screen "Lists" 1920x1080, template "Tpl"
   TextField "frm_1" at 16,154 size 1888x84; Text 'Text'
   TextField "txt_1" at 28,158 size 400x28; Text 'POSTAVKE (dok sustav stoji)'
   TextField "txt_2" at 28,194 size 160x34; Text 'Redoslijed'
   SymbolicIOField "sym_1" at 188,194 size 330x34; TextOff '0'; TextOn '1'; TextList "TL_Order"
      ProcessValue <- "CfgOrderMode"
   TextField "txt_3" at 560,194 size 290x34; Text 'SEMI: transfer po koraku'
   SymbolicIOField "sym_2" at 850,194 size 110x34; TextOff '0'; TextOn '1'; TextList "TL_YesNo"
      ProcessValue <- "CfgSemiPerTransfer"
   TextField "txt_4" at 1000,194 size 180x34; Text 'Ravnoteža'
   SymbolicIOField "sym_3" at 1180,194 size 260x34; TextOff '0'; TextOn '1'; TextList "TL_BalMode"
      ProcessValue <- "CfgBalMode"
   TextField "txt_5" at 1480,194 size 80x34; Text 'Istovar'
   IOField "io_1" at 1560,194 size 60x34; FormatPattern 99
      ProcessValue <- "UTotal"
   TextField "txt_6" at 1640,194 size 80x34; Text 'Ukrcaj'
   IOField "io_2" at 1720,194 size 60x34; FormatPattern 99
      ProcessValue <- "LTotal"
   TextField "txt_7" at 16,252 size 466x28; Text 'LISTA ZA ISTOVAR (DB20) 1-24'
   TextField "txt_8" at 16,286 size 46x27; Text '1'
   IOField "io_3" at 68,286 size 90x27; FormatPattern 999
      ProcessValue <- "UList_01"
   SymbolicIOField "sym_4" at 164,286 size 150x27; TextOff '0'; TextOn '1'; TextList "TL_ListSt"
      ProcessValue <- "UState_01"
   TextField "txt_9" at 16,316 size 46x27; Text '2'
   IOField "io_4" at 68,316 size 90x27; FormatPattern 999
      ProcessValue <- "UList_02"
   SymbolicIOField "sym_5" at 164,316 size 150x27; TextOff '0'; TextOn '1'; TextList "TL_ListSt"
      ProcessValue <- "UState_02"
   TextField "txt_10" at 16,346 size 46x27; Text '3'
   IOField "io_5" at 68,346 size 90x27; FormatPattern 999
      ProcessValue <- "UList_03"
   SymbolicIOField "sym_6" at 164,346 size 150x27; TextOff '0'; TextOn '1'; TextList "TL_ListSt"
      ProcessValue <- "UState_03"
   TextField "txt_11" at 16,376 size 46x27; Text '4'
   IOField "io_6" at 68,376 size 90x27; FormatPattern 999
      ProcessValue <- "UList_04"
   SymbolicIOField "sym_7" at 164,376 size 150x27; TextOff '0'; TextOn '1'; TextList "TL_ListSt"
      ProcessValue <- "UState_04"
   TextField "txt_12" at 16,406 size 46x27; Text '5'
   IOField "io_7" at 68,406 size 90x27; FormatPattern 999
      ProcessValue <- "UList_05"
   SymbolicIOField "sym_8" at 164,406 size 150x27; TextOff '0'; TextOn '1'; TextList "TL_ListSt"
      ProcessValue <- "UState_05"
   TextField "txt_13" at 16,436 size 46x27; Text '6'
   IOField "io_8" at 68,436 size 90x27; FormatPattern 999
      ProcessValue <- "UList_06"
   SymbolicIOField "sym_9" at 164,436 size 150x27; TextOff '0'; TextOn '1'; TextList "TL_ListSt"
      ProcessValue <- "UState_06"
   TextField "txt_14" at 16,466 size 46x27; Text '7'
   IOField "io_9" at 68,466 size 90x27; FormatPattern 999
      ProcessValue <- "UList_07"
   SymbolicIOField "sym_10" at 164,466 size 150x27; TextOff '0'; TextOn '1'; TextList "TL_ListSt"
      ProcessValue <- "UState_07"
   TextField "txt_15" at 16,496 size 46x27; Text '8'
   IOField "io_10" at 68,496 size 90x27; FormatPattern 999
      ProcessValue <- "UList_08"
   SymbolicIOField "sym_11" at 164,496 size 150x27; TextOff '0'; TextOn '1'; TextList "TL_ListSt"
      ProcessValue <- "UState_08"
   TextField "txt_16" at 16,526 size 46x27; Text '9'
   IOField "io_11" at 68,526 size 90x27; FormatPattern 999
      ProcessValue <- "UList_09"
   SymbolicIOField "sym_12" at 164,526 size 150x27; TextOff '0'; TextOn '1'; TextList "TL_ListSt"
      ProcessValue <- "UState_09"
   TextField "txt_17" at 16,556 size 46x27; Text '10'
   IOField "io_12" at 68,556 size 90x27; FormatPattern 999
      ProcessValue <- "UList_10"
   SymbolicIOField "sym_13" at 164,556 size 150x27; TextOff '0'; TextOn '1'; TextList "TL_ListSt"
      ProcessValue <- "UState_10"
   TextField "txt_18" at 16,586 size 46x27; Text '11'
   IOField "io_13" at 68,586 size 90x27; FormatPattern 999
      ProcessValue <- "UList_11"
   SymbolicIOField "sym_14" at 164,586 size 150x27; TextOff '0'; TextOn '1'; TextList "TL_ListSt"
      ProcessValue <- "UState_11"
   TextField "txt_19" at 16,616 size 46x27; Text '12'
   IOField "io_14" at 68,616 size 90x27; FormatPattern 999
      ProcessValue <- "UList_12"
   SymbolicIOField "sym_15" at 164,616 size 150x27; TextOff '0'; TextOn '1'; TextList "TL_ListSt"
      ProcessValue <- "UState_12"
   TextField "txt_20" at 16,646 size 46x27; Text '13'
   IOField "io_15" at 68,646 size 90x27; FormatPattern 999
      ProcessValue <- "UList_13"
   SymbolicIOField "sym_16" at 164,646 size 150x27; TextOff '0'; TextOn '1'; TextList "TL_ListSt"
      ProcessValue <- "UState_13"
   TextField "txt_21" at 16,676 size 46x27; Text '14'
   IOField "io_16" at 68,676 size 90x27; FormatPattern 999
      ProcessValue <- "UList_14"
   SymbolicIOField "sym_17" at 164,676 size 150x27; TextOff '0'; TextOn '1'; TextList "TL_ListSt"
      ProcessValue <- "UState_14"
   TextField "txt_22" at 16,706 size 46x27; Text '15'
   IOField "io_17" at 68,706 size 90x27; FormatPattern 999
      ProcessValue <- "UList_15"
   SymbolicIOField "sym_18" at 164,706 size 150x27; TextOff '0'; TextOn '1'; TextList "TL_ListSt"
      ProcessValue <- "UState_15"
   TextField "txt_23" at 16,736 size 46x27; Text '16'
   IOField "io_18" at 68,736 size 90x27; FormatPattern 999
      ProcessValue <- "UList_16"
   SymbolicIOField "sym_19" at 164,736 size 150x27; TextOff '0'; TextOn '1'; TextList "TL_ListSt"
      ProcessValue <- "UState_16"
   TextField "txt_24" at 16,766 size 46x27; Text '17'
   IOField "io_19" at 68,766 size 90x27; FormatPattern 999
      ProcessValue <- "UList_17"
   SymbolicIOField "sym_20" at 164,766 size 150x27; TextOff '0'; TextOn '1'; TextList "TL_ListSt"
      ProcessValue <- "UState_17"
   TextField "txt_25" at 16,796 size 46x27; Text '18'
   IOField "io_20" at 68,796 size 90x27; FormatPattern 999
      ProcessValue <- "UList_18"
   SymbolicIOField "sym_21" at 164,796 size 150x27; TextOff '0'; TextOn '1'; TextList "TL_ListSt"
      ProcessValue <- "UState_18"
   TextField "txt_26" at 16,826 size 46x27; Text '19'
   IOField "io_21" at 68,826 size 90x27; FormatPattern 999
      ProcessValue <- "UList_19"
   SymbolicIOField "sym_22" at 164,826 size 150x27; TextOff '0'; TextOn '1'; TextList "TL_ListSt"
      ProcessValue <- "UState_19"
   TextField "txt_27" at 16,856 size 46x27; Text '20'
   IOField "io_22" at 68,856 size 90x27; FormatPattern 999
      ProcessValue <- "UList_20"
   SymbolicIOField "sym_23" at 164,856 size 150x27; TextOff '0'; TextOn '1'; TextList "TL_ListSt"
      ProcessValue <- "UState_20"
   TextField "txt_28" at 16,886 size 46x27; Text '21'
   IOField "io_23" at 68,886 size 90x27; FormatPattern 999
      ProcessValue <- "UList_21"
   SymbolicIOField "sym_24" at 164,886 size 150x27; TextOff '0'; TextOn '1'; TextList "TL_ListSt"
      ProcessValue <- "UState_21"
   TextField "txt_29" at 16,916 size 46x27; Text '22'
   IOField "io_24" at 68,916 size 90x27; FormatPattern 999
      ProcessValue <- "UList_22"
   SymbolicIOField "sym_25" at 164,916 size 150x27; TextOff '0'; TextOn '1'; TextList "TL_ListSt"
      ProcessValue <- "UState_22"
   TextField "txt_30" at 16,946 size 46x27; Text '23'
   IOField "io_25" at 68,946 size 90x27; FormatPattern 999
      ProcessValue <- "UList_23"
   SymbolicIOField "sym_26" at 164,946 size 150x27; TextOff '0'; TextOn '1'; TextList "TL_ListSt"
      ProcessValue <- "UState_23"
   TextField "txt_31" at 16,976 size 46x27; Text '24'
   IOField "io_26" at 68,976 size 90x27; FormatPattern 999
      ProcessValue <- "UList_24"
   SymbolicIOField "sym_27" at 164,976 size 150x27; TextOff '0'; TextOn '1'; TextList "TL_ListSt"
      ProcessValue <- "UState_24"
   TextField "txt_32" at 490,252 size 466x28; Text 'LISTA ZA ISTOVAR 25-48'
   TextField "txt_33" at 490,286 size 46x27; Text '25'
   IOField "io_27" at 542,286 size 90x27; FormatPattern 999
      ProcessValue <- "UList_25"
   SymbolicIOField "sym_28" at 638,286 size 150x27; TextOff '0'; TextOn '1'; TextList "TL_ListSt"
      ProcessValue <- "UState_25"
   TextField "txt_34" at 490,316 size 46x27; Text '26'
   IOField "io_28" at 542,316 size 90x27; FormatPattern 999
      ProcessValue <- "UList_26"
   SymbolicIOField "sym_29" at 638,316 size 150x27; TextOff '0'; TextOn '1'; TextList "TL_ListSt"
      ProcessValue <- "UState_26"
   TextField "txt_35" at 490,346 size 46x27; Text '27'
   IOField "io_29" at 542,346 size 90x27; FormatPattern 999
      ProcessValue <- "UList_27"
   SymbolicIOField "sym_30" at 638,346 size 150x27; TextOff '0'; TextOn '1'; TextList "TL_ListSt"
      ProcessValue <- "UState_27"
   TextField "txt_36" at 490,376 size 46x27; Text '28'
   IOField "io_30" at 542,376 size 90x27; FormatPattern 999
      ProcessValue <- "UList_28"
   SymbolicIOField "sym_31" at 638,376 size 150x27; TextOff '0'; TextOn '1'; TextList "TL_ListSt"
      ProcessValue <- "UState_28"
   TextField "txt_37" at 490,406 size 46x27; Text '29'
   IOField "io_31" at 542,406 size 90x27; FormatPattern 999
      ProcessValue <- "UList_29"
   SymbolicIOField "sym_32" at 638,406 size 150x27; TextOff '0'; TextOn '1'; TextList "TL_ListSt"
      ProcessValue <- "UState_29"
   TextField "txt_38" at 490,436 size 46x27; Text '30'
   IOField "io_32" at 542,436 size 90x27; FormatPattern 999
      ProcessValue <- "UList_30"
   SymbolicIOField "sym_33" at 638,436 size 150x27; TextOff '0'; TextOn '1'; TextList "TL_ListSt"
      ProcessValue <- "UState_30"
   TextField "txt_39" at 490,466 size 46x27; Text '31'
   IOField "io_33" at 542,466 size 90x27; FormatPattern 999
      ProcessValue <- "UList_31"
   SymbolicIOField "sym_34" at 638,466 size 150x27; TextOff '0'; TextOn '1'; TextList "TL_ListSt"
      ProcessValue <- "UState_31"
   TextField "txt_40" at 490,496 size 46x27; Text '32'
   IOField "io_34" at 542,496 size 90x27; FormatPattern 999
      ProcessValue <- "UList_32"
   SymbolicIOField "sym_35" at 638,496 size 150x27; TextOff '0'; TextOn '1'; TextList "TL_ListSt"
      ProcessValue <- "UState_32"
   TextField "txt_41" at 490,526 size 46x27; Text '33'
   IOField "io_35" at 542,526 size 90x27; FormatPattern 999
      ProcessValue <- "UList_33"
   SymbolicIOField "sym_36" at 638,526 size 150x27; TextOff '0'; TextOn '1'; TextList "TL_ListSt"
      ProcessValue <- "UState_33"
   TextField "txt_42" at 490,556 size 46x27; Text '34'
   IOField "io_36" at 542,556 size 90x27; FormatPattern 999
      ProcessValue <- "UList_34"
   SymbolicIOField "sym_37" at 638,556 size 150x27; TextOff '0'; TextOn '1'; TextList "TL_ListSt"
      ProcessValue <- "UState_34"
   TextField "txt_43" at 490,586 size 46x27; Text '35'
   IOField "io_37" at 542,586 size 90x27; FormatPattern 999
      ProcessValue <- "UList_35"
   SymbolicIOField "sym_38" at 638,586 size 150x27; TextOff '0'; TextOn '1'; TextList "TL_ListSt"
      ProcessValue <- "UState_35"
   TextField "txt_44" at 490,616 size 46x27; Text '36'
   IOField "io_38" at 542,616 size 90x27; FormatPattern 999
      ProcessValue <- "UList_36"
   SymbolicIOField "sym_39" at 638,616 size 150x27; TextOff '0'; TextOn '1'; TextList "TL_ListSt"
      ProcessValue <- "UState_36"
   TextField "txt_45" at 490,646 size 46x27; Text '37'
   IOField "io_39" at 542,646 size 90x27; FormatPattern 999
      ProcessValue <- "UList_37"
   SymbolicIOField "sym_40" at 638,646 size 150x27; TextOff '0'; TextOn '1'; TextList "TL_ListSt"
      ProcessValue <- "UState_37"
   TextField "txt_46" at 490,676 size 46x27; Text '38'
   IOField "io_40" at 542,676 size 90x27; FormatPattern 999
      ProcessValue <- "UList_38"
   SymbolicIOField "sym_41" at 638,676 size 150x27; TextOff '0'; TextOn '1'; TextList "TL_ListSt"
      ProcessValue <- "UState_38"
   TextField "txt_47" at 490,706 size 46x27; Text '39'
   IOField "io_41" at 542,706 size 90x27; FormatPattern 999
      ProcessValue <- "UList_39"
   SymbolicIOField "sym_42" at 638,706 size 150x27; TextOff '0'; TextOn '1'; TextList "TL_ListSt"
      ProcessValue <- "UState_39"
   TextField "txt_48" at 490,736 size 46x27; Text '40'
   IOField "io_42" at 542,736 size 90x27; FormatPattern 999
      ProcessValue <- "UList_40"
   SymbolicIOField "sym_43" at 638,736 size 150x27; TextOff '0'; TextOn '1'; TextList "TL_ListSt"
      ProcessValue <- "UState_40"
   TextField "txt_49" at 490,766 size 46x27; Text '41'
   IOField "io_43" at 542,766 size 90x27; FormatPattern 999
      ProcessValue <- "UList_41"
   SymbolicIOField "sym_44" at 638,766 size 150x27; TextOff '0'; TextOn '1'; TextList "TL_ListSt"
      ProcessValue <- "UState_41"
   TextField "txt_50" at 490,796 size 46x27; Text '42'
   IOField "io_44" at 542,796 size 90x27; FormatPattern 999
      ProcessValue <- "UList_42"
   SymbolicIOField "sym_45" at 638,796 size 150x27; TextOff '0'; TextOn '1'; TextList "TL_ListSt"
      ProcessValue <- "UState_42"
   TextField "txt_51" at 490,826 size 46x27; Text '43'
   IOField "io_45" at 542,826 size 90x27; FormatPattern 999
      ProcessValue <- "UList_43"
   SymbolicIOField "sym_46" at 638,826 size 150x27; TextOff '0'; TextOn '1'; TextList "TL_ListSt"
      ProcessValue <- "UState_43"
   TextField "txt_52" at 490,856 size 46x27; Text '44'
   IOField "io_46" at 542,856 size 90x27; FormatPattern 999
      ProcessValue <- "UList_44"
   SymbolicIOField "sym_47" at 638,856 size 150x27; TextOff '0'; TextOn '1'; TextList "TL_ListSt"
      ProcessValue <- "UState_44"
   TextField "txt_53" at 490,886 size 46x27; Text '45'
   IOField "io_47" at 542,886 size 90x27; FormatPattern 999
      ProcessValue <- "UList_45"
   SymbolicIOField "sym_48" at 638,886 size 150x27; TextOff '0'; TextOn '1'; TextList "TL_ListSt"
      ProcessValue <- "UState_45"
   TextField "txt_54" at 490,916 size 46x27; Text '46'
   IOField "io_48" at 542,916 size 90x27; FormatPattern 999
      ProcessValue <- "UList_46"
   SymbolicIOField "sym_49" at 638,916 size 150x27; TextOff '0'; TextOn '1'; TextList "TL_ListSt"
      ProcessValue <- "UState_46"
   TextField "txt_55" at 490,946 size 46x27; Text '47'
   IOField "io_49" at 542,946 size 90x27; FormatPattern 999
      ProcessValue <- "UList_47"
   SymbolicIOField "sym_50" at 638,946 size 150x27; TextOff '0'; TextOn '1'; TextList "TL_ListSt"
      ProcessValue <- "UState_47"
   TextField "txt_56" at 490,976 size 46x27; Text '48'
   IOField "io_50" at 542,976 size 90x27; FormatPattern 999
      ProcessValue <- "UList_48"
   SymbolicIOField "sym_51" at 638,976 size 150x27; TextOff '0'; TextOn '1'; TextList "TL_ListSt"
      ProcessValue <- "UState_48"
   TextField "txt_57" at 964,252 size 466x28; Text 'LISTA ZA UKRCAJ (DB21) 1-24'
   TextField "txt_58" at 964,286 size 46x27; Text '1'
   IOField "io_51" at 1016,286 size 90x27; FormatPattern 999
      ProcessValue <- "LList_01"
   SymbolicIOField "sym_52" at 1112,286 size 150x27; TextOff '0'; TextOn '1'; TextList "TL_ListSt"
      ProcessValue <- "LState_01"
   TextField "txt_59" at 964,316 size 46x27; Text '2'
   IOField "io_52" at 1016,316 size 90x27; FormatPattern 999
      ProcessValue <- "LList_02"
   SymbolicIOField "sym_53" at 1112,316 size 150x27; TextOff '0'; TextOn '1'; TextList "TL_ListSt"
      ProcessValue <- "LState_02"
   TextField "txt_60" at 964,346 size 46x27; Text '3'
   IOField "io_53" at 1016,346 size 90x27; FormatPattern 999
      ProcessValue <- "LList_03"
   SymbolicIOField "sym_54" at 1112,346 size 150x27; TextOff '0'; TextOn '1'; TextList "TL_ListSt"
      ProcessValue <- "LState_03"
   TextField "txt_61" at 964,376 size 46x27; Text '4'
   IOField "io_54" at 1016,376 size 90x27; FormatPattern 999
      ProcessValue <- "LList_04"
   SymbolicIOField "sym_55" at 1112,376 size 150x27; TextOff '0'; TextOn '1'; TextList "TL_ListSt"
      ProcessValue <- "LState_04"
   TextField "txt_62" at 964,406 size 46x27; Text '5'
   IOField "io_55" at 1016,406 size 90x27; FormatPattern 999
      ProcessValue <- "LList_05"
   SymbolicIOField "sym_56" at 1112,406 size 150x27; TextOff '0'; TextOn '1'; TextList "TL_ListSt"
      ProcessValue <- "LState_05"
   TextField "txt_63" at 964,436 size 46x27; Text '6'
   IOField "io_56" at 1016,436 size 90x27; FormatPattern 999
      ProcessValue <- "LList_06"
   SymbolicIOField "sym_57" at 1112,436 size 150x27; TextOff '0'; TextOn '1'; TextList "TL_ListSt"
      ProcessValue <- "LState_06"
   TextField "txt_64" at 964,466 size 46x27; Text '7'
   IOField "io_57" at 1016,466 size 90x27; FormatPattern 999
      ProcessValue <- "LList_07"
   SymbolicIOField "sym_58" at 1112,466 size 150x27; TextOff '0'; TextOn '1'; TextList "TL_ListSt"
      ProcessValue <- "LState_07"
   TextField "txt_65" at 964,496 size 46x27; Text '8'
   IOField "io_58" at 1016,496 size 90x27; FormatPattern 999
      ProcessValue <- "LList_08"
   SymbolicIOField "sym_59" at 1112,496 size 150x27; TextOff '0'; TextOn '1'; TextList "TL_ListSt"
      ProcessValue <- "LState_08"
   TextField "txt_66" at 964,526 size 46x27; Text '9'
   IOField "io_59" at 1016,526 size 90x27; FormatPattern 999
      ProcessValue <- "LList_09"
   SymbolicIOField "sym_60" at 1112,526 size 150x27; TextOff '0'; TextOn '1'; TextList "TL_ListSt"
      ProcessValue <- "LState_09"
   TextField "txt_67" at 964,556 size 46x27; Text '10'
   IOField "io_60" at 1016,556 size 90x27; FormatPattern 999
      ProcessValue <- "LList_10"
   SymbolicIOField "sym_61" at 1112,556 size 150x27; TextOff '0'; TextOn '1'; TextList "TL_ListSt"
      ProcessValue <- "LState_10"
   TextField "txt_68" at 964,586 size 46x27; Text '11'
   IOField "io_61" at 1016,586 size 90x27; FormatPattern 999
      ProcessValue <- "LList_11"
   SymbolicIOField "sym_62" at 1112,586 size 150x27; TextOff '0'; TextOn '1'; TextList "TL_ListSt"
      ProcessValue <- "LState_11"
   TextField "txt_69" at 964,616 size 46x27; Text '12'
   IOField "io_62" at 1016,616 size 90x27; FormatPattern 999
      ProcessValue <- "LList_12"
   SymbolicIOField "sym_63" at 1112,616 size 150x27; TextOff '0'; TextOn '1'; TextList "TL_ListSt"
      ProcessValue <- "LState_12"
   TextField "txt_70" at 964,646 size 46x27; Text '13'
   IOField "io_63" at 1016,646 size 90x27; FormatPattern 999
      ProcessValue <- "LList_13"
   SymbolicIOField "sym_64" at 1112,646 size 150x27; TextOff '0'; TextOn '1'; TextList "TL_ListSt"
      ProcessValue <- "LState_13"
   TextField "txt_71" at 964,676 size 46x27; Text '14'
   IOField "io_64" at 1016,676 size 90x27; FormatPattern 999
      ProcessValue <- "LList_14"
   SymbolicIOField "sym_65" at 1112,676 size 150x27; TextOff '0'; TextOn '1'; TextList "TL_ListSt"
      ProcessValue <- "LState_14"
   TextField "txt_72" at 964,706 size 46x27; Text '15'
   IOField "io_65" at 1016,706 size 90x27; FormatPattern 999
      ProcessValue <- "LList_15"
   SymbolicIOField "sym_66" at 1112,706 size 150x27; TextOff '0'; TextOn '1'; TextList "TL_ListSt"
      ProcessValue <- "LState_15"
   TextField "txt_73" at 964,736 size 46x27; Text '16'
   IOField "io_66" at 1016,736 size 90x27; FormatPattern 999
      ProcessValue <- "LList_16"
   SymbolicIOField "sym_67" at 1112,736 size 150x27; TextOff '0'; TextOn '1'; TextList "TL_ListSt"
      ProcessValue <- "LState_16"
   TextField "txt_74" at 964,766 size 46x27; Text '17'
   IOField "io_67" at 1016,766 size 90x27; FormatPattern 999
      ProcessValue <- "LList_17"
   SymbolicIOField "sym_68" at 1112,766 size 150x27; TextOff '0'; TextOn '1'; TextList "TL_ListSt"
      ProcessValue <- "LState_17"
   TextField "txt_75" at 964,796 size 46x27; Text '18'
   IOField "io_68" at 1016,796 size 90x27; FormatPattern 999
      ProcessValue <- "LList_18"
   SymbolicIOField "sym_69" at 1112,796 size 150x27; TextOff '0'; TextOn '1'; TextList "TL_ListSt"
      ProcessValue <- "LState_18"
   TextField "txt_76" at 964,826 size 46x27; Text '19'
   IOField "io_69" at 1016,826 size 90x27; FormatPattern 999
      ProcessValue <- "LList_19"
   SymbolicIOField "sym_70" at 1112,826 size 150x27; TextOff '0'; TextOn '1'; TextList "TL_ListSt"
      ProcessValue <- "LState_19"
   TextField "txt_77" at 964,856 size 46x27; Text '20'
   IOField "io_70" at 1016,856 size 90x27; FormatPattern 999
      ProcessValue <- "LList_20"
   SymbolicIOField "sym_71" at 1112,856 size 150x27; TextOff '0'; TextOn '1'; TextList "TL_ListSt"
      ProcessValue <- "LState_20"
   TextField "txt_78" at 964,886 size 46x27; Text '21'
   IOField "io_71" at 1016,886 size 90x27; FormatPattern 999
      ProcessValue <- "LList_21"
   SymbolicIOField "sym_72" at 1112,886 size 150x27; TextOff '0'; TextOn '1'; TextList "TL_ListSt"
      ProcessValue <- "LState_21"
   TextField "txt_79" at 964,916 size 46x27; Text '22'
   IOField "io_72" at 1016,916 size 90x27; FormatPattern 999
      ProcessValue <- "LList_22"
   SymbolicIOField "sym_73" at 1112,916 size 150x27; TextOff '0'; TextOn '1'; TextList "TL_ListSt"
      ProcessValue <- "LState_22"
   TextField "txt_80" at 964,946 size 46x27; Text '23'
   IOField "io_73" at 1016,946 size 90x27; FormatPattern 999
      ProcessValue <- "LList_23"
   SymbolicIOField "sym_74" at 1112,946 size 150x27; TextOff '0'; TextOn '1'; TextList "TL_ListSt"
      ProcessValue <- "LState_23"
   TextField "txt_81" at 964,976 size 46x27; Text '24'
   IOField "io_74" at 1016,976 size 90x27; FormatPattern 999
      ProcessValue <- "LList_24"
   SymbolicIOField "sym_75" at 1112,976 size 150x27; TextOff '0'; TextOn '1'; TextList "TL_ListSt"
      ProcessValue <- "LState_24"
   TextField "txt_82" at 1438,252 size 466x28; Text 'LISTA ZA UKRCAJ 25-48'
   TextField "txt_83" at 1438,286 size 46x27; Text '25'
   IOField "io_75" at 1490,286 size 90x27; FormatPattern 999
      ProcessValue <- "LList_25"
   SymbolicIOField "sym_76" at 1586,286 size 150x27; TextOff '0'; TextOn '1'; TextList "TL_ListSt"
      ProcessValue <- "LState_25"
   TextField "txt_84" at 1438,316 size 46x27; Text '26'
   IOField "io_76" at 1490,316 size 90x27; FormatPattern 999
      ProcessValue <- "LList_26"
   SymbolicIOField "sym_77" at 1586,316 size 150x27; TextOff '0'; TextOn '1'; TextList "TL_ListSt"
      ProcessValue <- "LState_26"
   TextField "txt_85" at 1438,346 size 46x27; Text '27'
   IOField "io_77" at 1490,346 size 90x27; FormatPattern 999
      ProcessValue <- "LList_27"
   SymbolicIOField "sym_78" at 1586,346 size 150x27; TextOff '0'; TextOn '1'; TextList "TL_ListSt"
      ProcessValue <- "LState_27"
   TextField "txt_86" at 1438,376 size 46x27; Text '28'
   IOField "io_78" at 1490,376 size 90x27; FormatPattern 999
      ProcessValue <- "LList_28"
   SymbolicIOField "sym_79" at 1586,376 size 150x27; TextOff '0'; TextOn '1'; TextList "TL_ListSt"
      ProcessValue <- "LState_28"
   TextField "txt_87" at 1438,406 size 46x27; Text '29'
   IOField "io_79" at 1490,406 size 90x27; FormatPattern 999
      ProcessValue <- "LList_29"
   SymbolicIOField "sym_80" at 1586,406 size 150x27; TextOff '0'; TextOn '1'; TextList "TL_ListSt"
      ProcessValue <- "LState_29"
   TextField "txt_88" at 1438,436 size 46x27; Text '30'
   IOField "io_80" at 1490,436 size 90x27; FormatPattern 999
      ProcessValue <- "LList_30"
   SymbolicIOField "sym_81" at 1586,436 size 150x27; TextOff '0'; TextOn '1'; TextList "TL_ListSt"
      ProcessValue <- "LState_30"
   TextField "txt_89" at 1438,466 size 46x27; Text '31'
   IOField "io_81" at 1490,466 size 90x27; FormatPattern 999
      ProcessValue <- "LList_31"
   SymbolicIOField "sym_82" at 1586,466 size 150x27; TextOff '0'; TextOn '1'; TextList "TL_ListSt"
      ProcessValue <- "LState_31"
   TextField "txt_90" at 1438,496 size 46x27; Text '32'
   IOField "io_82" at 1490,496 size 90x27; FormatPattern 999
      ProcessValue <- "LList_32"
   SymbolicIOField "sym_83" at 1586,496 size 150x27; TextOff '0'; TextOn '1'; TextList "TL_ListSt"
      ProcessValue <- "LState_32"
   TextField "txt_91" at 1438,526 size 46x27; Text '33'
   IOField "io_83" at 1490,526 size 90x27; FormatPattern 999
      ProcessValue <- "LList_33"
   SymbolicIOField "sym_84" at 1586,526 size 150x27; TextOff '0'; TextOn '1'; TextList "TL_ListSt"
      ProcessValue <- "LState_33"
   TextField "txt_92" at 1438,556 size 46x27; Text '34'
   IOField "io_84" at 1490,556 size 90x27; FormatPattern 999
      ProcessValue <- "LList_34"
   SymbolicIOField "sym_85" at 1586,556 size 150x27; TextOff '0'; TextOn '1'; TextList "TL_ListSt"
      ProcessValue <- "LState_34"
   TextField "txt_93" at 1438,586 size 46x27; Text '35'
   IOField "io_85" at 1490,586 size 90x27; FormatPattern 999
      ProcessValue <- "LList_35"
   SymbolicIOField "sym_86" at 1586,586 size 150x27; TextOff '0'; TextOn '1'; TextList "TL_ListSt"
      ProcessValue <- "LState_35"
   TextField "txt_94" at 1438,616 size 46x27; Text '36'
   IOField "io_86" at 1490,616 size 90x27; FormatPattern 999
      ProcessValue <- "LList_36"
   SymbolicIOField "sym_87" at 1586,616 size 150x27; TextOff '0'; TextOn '1'; TextList "TL_ListSt"
      ProcessValue <- "LState_36"
   TextField "txt_95" at 1438,646 size 46x27; Text '37'
   IOField "io_87" at 1490,646 size 90x27; FormatPattern 999
      ProcessValue <- "LList_37"
   SymbolicIOField "sym_88" at 1586,646 size 150x27; TextOff '0'; TextOn '1'; TextList "TL_ListSt"
      ProcessValue <- "LState_37"
   TextField "txt_96" at 1438,676 size 46x27; Text '38'
   IOField "io_88" at 1490,676 size 90x27; FormatPattern 999
      ProcessValue <- "LList_38"
   SymbolicIOField "sym_89" at 1586,676 size 150x27; TextOff '0'; TextOn '1'; TextList "TL_ListSt"
      ProcessValue <- "LState_38"
   TextField "txt_97" at 1438,706 size 46x27; Text '39'
   IOField "io_89" at 1490,706 size 90x27; FormatPattern 999
      ProcessValue <- "LList_39"
   SymbolicIOField "sym_90" at 1586,706 size 150x27; TextOff '0'; TextOn '1'; TextList "TL_ListSt"
      ProcessValue <- "LState_39"
   TextField "txt_98" at 1438,736 size 46x27; Text '40'
   IOField "io_90" at 1490,736 size 90x27; FormatPattern 999
      ProcessValue <- "LList_40"
   SymbolicIOField "sym_91" at 1586,736 size 150x27; TextOff '0'; TextOn '1'; TextList "TL_ListSt"
      ProcessValue <- "LState_40"
   TextField "txt_99" at 1438,766 size 46x27; Text '41'
   IOField "io_91" at 1490,766 size 90x27; FormatPattern 999
      ProcessValue <- "LList_41"
   SymbolicIOField "sym_92" at 1586,766 size 150x27; TextOff '0'; TextOn '1'; TextList "TL_ListSt"
      ProcessValue <- "LState_41"
   TextField "txt_100" at 1438,796 size 46x27; Text '42'
   IOField "io_92" at 1490,796 size 90x27; FormatPattern 999
      ProcessValue <- "LList_42"
   SymbolicIOField "sym_93" at 1586,796 size 150x27; TextOff '0'; TextOn '1'; TextList "TL_ListSt"
      ProcessValue <- "LState_42"
   TextField "txt_101" at 1438,826 size 46x27; Text '43'
   IOField "io_93" at 1490,826 size 90x27; FormatPattern 999
      ProcessValue <- "LList_43"
   SymbolicIOField "sym_94" at 1586,826 size 150x27; TextOff '0'; TextOn '1'; TextList "TL_ListSt"
      ProcessValue <- "LState_43"
   TextField "txt_102" at 1438,856 size 46x27; Text '44'
   IOField "io_94" at 1490,856 size 90x27; FormatPattern 999
      ProcessValue <- "LList_44"
   SymbolicIOField "sym_95" at 1586,856 size 150x27; TextOff '0'; TextOn '1'; TextList "TL_ListSt"
      ProcessValue <- "LState_44"
   TextField "txt_103" at 1438,886 size 46x27; Text '45'
   IOField "io_95" at 1490,886 size 90x27; FormatPattern 999
      ProcessValue <- "LList_45"
   SymbolicIOField "sym_96" at 1586,886 size 150x27; TextOff '0'; TextOn '1'; TextList "TL_ListSt"
      ProcessValue <- "LState_45"
   TextField "txt_104" at 1438,916 size 46x27; Text '46'
   IOField "io_96" at 1490,916 size 90x27; FormatPattern 999
      ProcessValue <- "LList_46"
   SymbolicIOField "sym_97" at 1586,916 size 150x27; TextOff '0'; TextOn '1'; TextList "TL_ListSt"
      ProcessValue <- "LState_46"
   TextField "txt_105" at 1438,946 size 46x27; Text '47'
   IOField "io_97" at 1490,946 size 90x27; FormatPattern 999
      ProcessValue <- "LList_47"
   SymbolicIOField "sym_98" at 1586,946 size 150x27; TextOff '0'; TextOn '1'; TextList "TL_ListSt"
      ProcessValue <- "LState_47"
   TextField "txt_106" at 1438,976 size 46x27; Text '48'
   IOField "io_98" at 1490,976 size 90x27; FormatPattern 999
      ProcessValue <- "LList_48"
   SymbolicIOField "sym_99" at 1586,976 size 150x27; TextOff '0'; TextOn '1'; TextList "TL_ListSt"
      ProcessValue <- "LState_48"

screen "Manual" 1920x1080, template "Tpl"
   TextField "txt_1" at 60,154 size 446x28; Text 'BAY 1 - SKLADIŠTE (yard)'
   TextField "txt_2" at 744,154 size 446x28; Text 'BAY 0 - BROD (ship)'
   TextField "frm_1" at 56,186 size 1138x36; Text 'Text'
   TextField "frm_2" at 556,224 size 140x722; Text 'Text'
   TextField "txt_3" at 556,950 size 140x22; Text 'OBALA / kran y'
   TextField "frm_3" at 52,220 size 462x730; Text 'Text'
   TextField "frm_4" at 736,220 size 462x730; Text 'Text'
   TextField "frm_5" at 965,220 size 4x730; Text 'Text'
   TextField "txt_4" at 16,244 size 40x22; Text 'y0'
   TextField "txt_5" at 16,304 size 40x22; Text 'y1'
   TextField "txt_6" at 16,364 size 40x22; Text 'y2'
   TextField "txt_7" at 16,424 size 40x22; Text 'y3'
   TextField "txt_8" at 16,484 size 40x22; Text 'y4'
   TextField "txt_9" at 16,544 size 40x22; Text 'y5'
   TextField "txt_10" at 16,604 size 40x22; Text 'y6'
   TextField "txt_11" at 16,664 size 40x22; Text 'y7'
   TextField "txt_12" at 16,724 size 40x22; Text 'y8'
   TextField "txt_13" at 16,784 size 40x22; Text 'y9'
   TextField "txt_14" at 16,844 size 40x22; Text 'y10'
   TextField "txt_15" at 16,904 size 40x22; Text 'y11'
   TextField "txt_16" at 60,952 size 104x20; Text 'x0'
   TextField "txt_17" at 174,952 size 104x20; Text 'x1'
   TextField "txt_18" at 288,952 size 104x20; Text 'x2'
   TextField "txt_19" at 402,952 size 104x20; Text 'x3'
   TextField "txt_20" at 744,952 size 104x20; Text 'x0'
   TextField "txt_21" at 858,952 size 104x20; Text 'x1'
   TextField "txt_22" at 972,952 size 104x20; Text 'x2'
   TextField "txt_23" at 1086,952 size 104x20; Text 'x3'
   TextField "txt_24" at 744,976 size 120x28; Text 'LIJEVO'
   IOField "io_1" at 864,976 size 60x28; FormatPattern 99
      ProcessValue <- "BalL"
   TextField "txt_25" at 972,976 size 120x28; Text 'DESNO'
   IOField "io_2" at 1092,976 size 60x28; FormatPattern 99
      ProcessValue <- "BalR"
   Rectangle "cel_1" at 60,228 size 104x54
      Appearance <- "CellSt1_00"
   IOField "io_3" at 67,235 size 90x40; FormatPattern 999
      ProcessValue <- "Cell1_00"
      Appearance <- "CellSt1_00"
   Rectangle "cel_2" at 60,288 size 104x54
      Appearance <- "CellSt1_01"
   IOField "io_4" at 67,295 size 90x40; FormatPattern 999
      ProcessValue <- "Cell1_01"
      Appearance <- "CellSt1_01"
   Rectangle "cel_3" at 60,348 size 104x54
      Appearance <- "CellSt1_02"
   IOField "io_5" at 67,355 size 90x40; FormatPattern 999
      ProcessValue <- "Cell1_02"
      Appearance <- "CellSt1_02"
   Rectangle "cel_4" at 60,408 size 104x54
      Appearance <- "CellSt1_03"
   IOField "io_6" at 67,415 size 90x40; FormatPattern 999
      ProcessValue <- "Cell1_03"
      Appearance <- "CellSt1_03"
   Rectangle "cel_5" at 60,468 size 104x54
      Appearance <- "CellSt1_04"
   IOField "io_7" at 67,475 size 90x40; FormatPattern 999
      ProcessValue <- "Cell1_04"
      Appearance <- "CellSt1_04"
   Rectangle "cel_6" at 60,528 size 104x54
      Appearance <- "CellSt1_05"
   IOField "io_8" at 67,535 size 90x40; FormatPattern 999
      ProcessValue <- "Cell1_05"
      Appearance <- "CellSt1_05"
   Rectangle "cel_7" at 60,588 size 104x54
      Appearance <- "CellSt1_06"
   IOField "io_9" at 67,595 size 90x40; FormatPattern 999
      ProcessValue <- "Cell1_06"
      Appearance <- "CellSt1_06"
   Rectangle "cel_8" at 60,648 size 104x54
      Appearance <- "CellSt1_07"
   IOField "io_10" at 67,655 size 90x40; FormatPattern 999
      ProcessValue <- "Cell1_07"
      Appearance <- "CellSt1_07"
   Rectangle "cel_9" at 60,708 size 104x54
      Appearance <- "CellSt1_08"
   IOField "io_11" at 67,715 size 90x40; FormatPattern 999
      ProcessValue <- "Cell1_08"
      Appearance <- "CellSt1_08"
   Rectangle "cel_10" at 60,768 size 104x54
      Appearance <- "CellSt1_09"
   IOField "io_12" at 67,775 size 90x40; FormatPattern 999
      ProcessValue <- "Cell1_09"
      Appearance <- "CellSt1_09"
   Rectangle "cel_11" at 60,828 size 104x54
      Appearance <- "CellSt1_10"
   IOField "io_13" at 67,835 size 90x40; FormatPattern 999
      ProcessValue <- "Cell1_10"
      Appearance <- "CellSt1_10"
   Rectangle "cel_12" at 60,888 size 104x54
      Appearance <- "CellSt1_11"
   IOField "io_14" at 67,895 size 90x40; FormatPattern 999
      ProcessValue <- "Cell1_11"
      Appearance <- "CellSt1_11"
   Rectangle "cel_13" at 174,228 size 104x54
      Appearance <- "CellSt1_12"
   IOField "io_15" at 181,235 size 90x40; FormatPattern 999
      ProcessValue <- "Cell1_12"
      Appearance <- "CellSt1_12"
   Rectangle "cel_14" at 174,288 size 104x54
      Appearance <- "CellSt1_13"
   IOField "io_16" at 181,295 size 90x40; FormatPattern 999
      ProcessValue <- "Cell1_13"
      Appearance <- "CellSt1_13"
   Rectangle "cel_15" at 174,348 size 104x54
      Appearance <- "CellSt1_14"
   IOField "io_17" at 181,355 size 90x40; FormatPattern 999
      ProcessValue <- "Cell1_14"
      Appearance <- "CellSt1_14"
   Rectangle "cel_16" at 174,408 size 104x54
      Appearance <- "CellSt1_15"
   IOField "io_18" at 181,415 size 90x40; FormatPattern 999
      ProcessValue <- "Cell1_15"
      Appearance <- "CellSt1_15"
   Rectangle "cel_17" at 174,468 size 104x54
      Appearance <- "CellSt1_16"
   IOField "io_19" at 181,475 size 90x40; FormatPattern 999
      ProcessValue <- "Cell1_16"
      Appearance <- "CellSt1_16"
   Rectangle "cel_18" at 174,528 size 104x54
      Appearance <- "CellSt1_17"
   IOField "io_20" at 181,535 size 90x40; FormatPattern 999
      ProcessValue <- "Cell1_17"
      Appearance <- "CellSt1_17"
   Rectangle "cel_19" at 174,588 size 104x54
      Appearance <- "CellSt1_18"
   IOField "io_21" at 181,595 size 90x40; FormatPattern 999
      ProcessValue <- "Cell1_18"
      Appearance <- "CellSt1_18"
   Rectangle "cel_20" at 174,648 size 104x54
      Appearance <- "CellSt1_19"
   IOField "io_22" at 181,655 size 90x40; FormatPattern 999
      ProcessValue <- "Cell1_19"
      Appearance <- "CellSt1_19"
   Rectangle "cel_21" at 174,708 size 104x54
      Appearance <- "CellSt1_20"
   IOField "io_23" at 181,715 size 90x40; FormatPattern 999
      ProcessValue <- "Cell1_20"
      Appearance <- "CellSt1_20"
   Rectangle "cel_22" at 174,768 size 104x54
      Appearance <- "CellSt1_21"
   IOField "io_24" at 181,775 size 90x40; FormatPattern 999
      ProcessValue <- "Cell1_21"
      Appearance <- "CellSt1_21"
   Rectangle "cel_23" at 174,828 size 104x54
      Appearance <- "CellSt1_22"
   IOField "io_25" at 181,835 size 90x40; FormatPattern 999
      ProcessValue <- "Cell1_22"
      Appearance <- "CellSt1_22"
   Rectangle "cel_24" at 174,888 size 104x54
      Appearance <- "CellSt1_23"
   IOField "io_26" at 181,895 size 90x40; FormatPattern 999
      ProcessValue <- "Cell1_23"
      Appearance <- "CellSt1_23"
   Rectangle "cel_25" at 288,228 size 104x54
      Appearance <- "CellSt1_24"
   IOField "io_27" at 295,235 size 90x40; FormatPattern 999
      ProcessValue <- "Cell1_24"
      Appearance <- "CellSt1_24"
   Rectangle "cel_26" at 288,288 size 104x54
      Appearance <- "CellSt1_25"
   IOField "io_28" at 295,295 size 90x40; FormatPattern 999
      ProcessValue <- "Cell1_25"
      Appearance <- "CellSt1_25"
   Rectangle "cel_27" at 288,348 size 104x54
      Appearance <- "CellSt1_26"
   IOField "io_29" at 295,355 size 90x40; FormatPattern 999
      ProcessValue <- "Cell1_26"
      Appearance <- "CellSt1_26"
   Rectangle "cel_28" at 288,408 size 104x54
      Appearance <- "CellSt1_27"
   IOField "io_30" at 295,415 size 90x40; FormatPattern 999
      ProcessValue <- "Cell1_27"
      Appearance <- "CellSt1_27"
   Rectangle "cel_29" at 288,468 size 104x54
      Appearance <- "CellSt1_28"
   IOField "io_31" at 295,475 size 90x40; FormatPattern 999
      ProcessValue <- "Cell1_28"
      Appearance <- "CellSt1_28"
   Rectangle "cel_30" at 288,528 size 104x54
      Appearance <- "CellSt1_29"
   IOField "io_32" at 295,535 size 90x40; FormatPattern 999
      ProcessValue <- "Cell1_29"
      Appearance <- "CellSt1_29"
   Rectangle "cel_31" at 288,588 size 104x54
      Appearance <- "CellSt1_30"
   IOField "io_33" at 295,595 size 90x40; FormatPattern 999
      ProcessValue <- "Cell1_30"
      Appearance <- "CellSt1_30"
   Rectangle "cel_32" at 288,648 size 104x54
      Appearance <- "CellSt1_31"
   IOField "io_34" at 295,655 size 90x40; FormatPattern 999
      ProcessValue <- "Cell1_31"
      Appearance <- "CellSt1_31"
   Rectangle "cel_33" at 288,708 size 104x54
      Appearance <- "CellSt1_32"
   IOField "io_35" at 295,715 size 90x40; FormatPattern 999
      ProcessValue <- "Cell1_32"
      Appearance <- "CellSt1_32"
   Rectangle "cel_34" at 288,768 size 104x54
      Appearance <- "CellSt1_33"
   IOField "io_36" at 295,775 size 90x40; FormatPattern 999
      ProcessValue <- "Cell1_33"
      Appearance <- "CellSt1_33"
   Rectangle "cel_35" at 288,828 size 104x54
      Appearance <- "CellSt1_34"
   IOField "io_37" at 295,835 size 90x40; FormatPattern 999
      ProcessValue <- "Cell1_34"
      Appearance <- "CellSt1_34"
   Rectangle "cel_36" at 288,888 size 104x54
      Appearance <- "CellSt1_35"
   IOField "io_38" at 295,895 size 90x40; FormatPattern 999
      ProcessValue <- "Cell1_35"
      Appearance <- "CellSt1_35"
   Rectangle "cel_37" at 402,228 size 104x54
      Appearance <- "CellSt1_36"
   IOField "io_39" at 409,235 size 90x40; FormatPattern 999
      ProcessValue <- "Cell1_36"
      Appearance <- "CellSt1_36"
   Rectangle "cel_38" at 402,288 size 104x54
      Appearance <- "CellSt1_37"
   IOField "io_40" at 409,295 size 90x40; FormatPattern 999
      ProcessValue <- "Cell1_37"
      Appearance <- "CellSt1_37"
   Rectangle "cel_39" at 402,348 size 104x54
      Appearance <- "CellSt1_38"
   IOField "io_41" at 409,355 size 90x40; FormatPattern 999
      ProcessValue <- "Cell1_38"
      Appearance <- "CellSt1_38"
   Rectangle "cel_40" at 402,408 size 104x54
      Appearance <- "CellSt1_39"
   IOField "io_42" at 409,415 size 90x40; FormatPattern 999
      ProcessValue <- "Cell1_39"
      Appearance <- "CellSt1_39"
   Rectangle "cel_41" at 402,468 size 104x54
      Appearance <- "CellSt1_40"
   IOField "io_43" at 409,475 size 90x40; FormatPattern 999
      ProcessValue <- "Cell1_40"
      Appearance <- "CellSt1_40"
   Rectangle "cel_42" at 402,528 size 104x54
      Appearance <- "CellSt1_41"
   IOField "io_44" at 409,535 size 90x40; FormatPattern 999
      ProcessValue <- "Cell1_41"
      Appearance <- "CellSt1_41"
   Rectangle "cel_43" at 402,588 size 104x54
      Appearance <- "CellSt1_42"
   IOField "io_45" at 409,595 size 90x40; FormatPattern 999
      ProcessValue <- "Cell1_42"
      Appearance <- "CellSt1_42"
   Rectangle "cel_44" at 402,648 size 104x54
      Appearance <- "CellSt1_43"
   IOField "io_46" at 409,655 size 90x40; FormatPattern 999
      ProcessValue <- "Cell1_43"
      Appearance <- "CellSt1_43"
   Rectangle "cel_45" at 402,708 size 104x54
      Appearance <- "CellSt1_44"
   IOField "io_47" at 409,715 size 90x40; FormatPattern 999
      ProcessValue <- "Cell1_44"
      Appearance <- "CellSt1_44"
   Rectangle "cel_46" at 402,768 size 104x54
      Appearance <- "CellSt1_45"
   IOField "io_48" at 409,775 size 90x40; FormatPattern 999
      ProcessValue <- "Cell1_45"
      Appearance <- "CellSt1_45"
   Rectangle "cel_47" at 402,828 size 104x54
      Appearance <- "CellSt1_46"
   IOField "io_49" at 409,835 size 90x40; FormatPattern 999
      ProcessValue <- "Cell1_46"
      Appearance <- "CellSt1_46"
   Rectangle "cel_48" at 402,888 size 104x54
      Appearance <- "CellSt1_47"
   IOField "io_50" at 409,895 size 90x40; FormatPattern 999
      ProcessValue <- "Cell1_47"
      Appearance <- "CellSt1_47"
   Rectangle "cel_49" at 744,228 size 104x54
      Appearance <- "CellSt0_00"
   IOField "io_51" at 751,235 size 90x40; FormatPattern 999
      ProcessValue <- "Cell0_00"
      Appearance <- "CellSt0_00"
   Rectangle "cel_50" at 744,288 size 104x54
      Appearance <- "CellSt0_01"
   IOField "io_52" at 751,295 size 90x40; FormatPattern 999
      ProcessValue <- "Cell0_01"
      Appearance <- "CellSt0_01"
   Rectangle "cel_51" at 744,348 size 104x54
      Appearance <- "CellSt0_02"
   IOField "io_53" at 751,355 size 90x40; FormatPattern 999
      ProcessValue <- "Cell0_02"
      Appearance <- "CellSt0_02"
   Rectangle "cel_52" at 744,408 size 104x54
      Appearance <- "CellSt0_03"
   IOField "io_54" at 751,415 size 90x40; FormatPattern 999
      ProcessValue <- "Cell0_03"
      Appearance <- "CellSt0_03"
   Rectangle "cel_53" at 744,468 size 104x54
      Appearance <- "CellSt0_04"
   IOField "io_55" at 751,475 size 90x40; FormatPattern 999
      ProcessValue <- "Cell0_04"
      Appearance <- "CellSt0_04"
   Rectangle "cel_54" at 744,528 size 104x54
      Appearance <- "CellSt0_05"
   IOField "io_56" at 751,535 size 90x40; FormatPattern 999
      ProcessValue <- "Cell0_05"
      Appearance <- "CellSt0_05"
   Rectangle "cel_55" at 744,588 size 104x54
      Appearance <- "CellSt0_06"
   IOField "io_57" at 751,595 size 90x40; FormatPattern 999
      ProcessValue <- "Cell0_06"
      Appearance <- "CellSt0_06"
   Rectangle "cel_56" at 744,648 size 104x54
      Appearance <- "CellSt0_07"
   IOField "io_58" at 751,655 size 90x40; FormatPattern 999
      ProcessValue <- "Cell0_07"
      Appearance <- "CellSt0_07"
   Rectangle "cel_57" at 744,708 size 104x54
      Appearance <- "CellSt0_08"
   IOField "io_59" at 751,715 size 90x40; FormatPattern 999
      ProcessValue <- "Cell0_08"
      Appearance <- "CellSt0_08"
   Rectangle "cel_58" at 744,768 size 104x54
      Appearance <- "CellSt0_09"
   IOField "io_60" at 751,775 size 90x40; FormatPattern 999
      ProcessValue <- "Cell0_09"
      Appearance <- "CellSt0_09"
   Rectangle "cel_59" at 744,828 size 104x54
      Appearance <- "CellSt0_10"
   IOField "io_61" at 751,835 size 90x40; FormatPattern 999
      ProcessValue <- "Cell0_10"
      Appearance <- "CellSt0_10"
   Rectangle "cel_60" at 744,888 size 104x54
      Appearance <- "CellSt0_11"
   IOField "io_62" at 751,895 size 90x40; FormatPattern 999
      ProcessValue <- "Cell0_11"
      Appearance <- "CellSt0_11"
   Rectangle "cel_61" at 858,228 size 104x54
      Appearance <- "CellSt0_12"
   IOField "io_63" at 865,235 size 90x40; FormatPattern 999
      ProcessValue <- "Cell0_12"
      Appearance <- "CellSt0_12"
   Rectangle "cel_62" at 858,288 size 104x54
      Appearance <- "CellSt0_13"
   IOField "io_64" at 865,295 size 90x40; FormatPattern 999
      ProcessValue <- "Cell0_13"
      Appearance <- "CellSt0_13"
   Rectangle "cel_63" at 858,348 size 104x54
      Appearance <- "CellSt0_14"
   IOField "io_65" at 865,355 size 90x40; FormatPattern 999
      ProcessValue <- "Cell0_14"
      Appearance <- "CellSt0_14"
   Rectangle "cel_64" at 858,408 size 104x54
      Appearance <- "CellSt0_15"
   IOField "io_66" at 865,415 size 90x40; FormatPattern 999
      ProcessValue <- "Cell0_15"
      Appearance <- "CellSt0_15"
   Rectangle "cel_65" at 858,468 size 104x54
      Appearance <- "CellSt0_16"
   IOField "io_67" at 865,475 size 90x40; FormatPattern 999
      ProcessValue <- "Cell0_16"
      Appearance <- "CellSt0_16"
   Rectangle "cel_66" at 858,528 size 104x54
      Appearance <- "CellSt0_17"
   IOField "io_68" at 865,535 size 90x40; FormatPattern 999
      ProcessValue <- "Cell0_17"
      Appearance <- "CellSt0_17"
   Rectangle "cel_67" at 858,588 size 104x54
      Appearance <- "CellSt0_18"
   IOField "io_69" at 865,595 size 90x40; FormatPattern 999
      ProcessValue <- "Cell0_18"
      Appearance <- "CellSt0_18"
   Rectangle "cel_68" at 858,648 size 104x54
      Appearance <- "CellSt0_19"
   IOField "io_70" at 865,655 size 90x40; FormatPattern 999
      ProcessValue <- "Cell0_19"
      Appearance <- "CellSt0_19"
   Rectangle "cel_69" at 858,708 size 104x54
      Appearance <- "CellSt0_20"
   IOField "io_71" at 865,715 size 90x40; FormatPattern 999
      ProcessValue <- "Cell0_20"
      Appearance <- "CellSt0_20"
   Rectangle "cel_70" at 858,768 size 104x54
      Appearance <- "CellSt0_21"
   IOField "io_72" at 865,775 size 90x40; FormatPattern 999
      ProcessValue <- "Cell0_21"
      Appearance <- "CellSt0_21"
   Rectangle "cel_71" at 858,828 size 104x54
      Appearance <- "CellSt0_22"
   IOField "io_73" at 865,835 size 90x40; FormatPattern 999
      ProcessValue <- "Cell0_22"
      Appearance <- "CellSt0_22"
   Rectangle "cel_72" at 858,888 size 104x54
      Appearance <- "CellSt0_23"
   IOField "io_74" at 865,895 size 90x40; FormatPattern 999
      ProcessValue <- "Cell0_23"
      Appearance <- "CellSt0_23"
   Rectangle "cel_73" at 972,228 size 104x54
      Appearance <- "CellSt0_24"
   IOField "io_75" at 979,235 size 90x40; FormatPattern 999
      ProcessValue <- "Cell0_24"
      Appearance <- "CellSt0_24"
   Rectangle "cel_74" at 972,288 size 104x54
      Appearance <- "CellSt0_25"
   IOField "io_76" at 979,295 size 90x40; FormatPattern 999
      ProcessValue <- "Cell0_25"
      Appearance <- "CellSt0_25"
   Rectangle "cel_75" at 972,348 size 104x54
      Appearance <- "CellSt0_26"
   IOField "io_77" at 979,355 size 90x40; FormatPattern 999
      ProcessValue <- "Cell0_26"
      Appearance <- "CellSt0_26"
   Rectangle "cel_76" at 972,408 size 104x54
      Appearance <- "CellSt0_27"
   IOField "io_78" at 979,415 size 90x40; FormatPattern 999
      ProcessValue <- "Cell0_27"
      Appearance <- "CellSt0_27"
   Rectangle "cel_77" at 972,468 size 104x54
      Appearance <- "CellSt0_28"
   IOField "io_79" at 979,475 size 90x40; FormatPattern 999
      ProcessValue <- "Cell0_28"
      Appearance <- "CellSt0_28"
   Rectangle "cel_78" at 972,528 size 104x54
      Appearance <- "CellSt0_29"
   IOField "io_80" at 979,535 size 90x40; FormatPattern 999
      ProcessValue <- "Cell0_29"
      Appearance <- "CellSt0_29"
   Rectangle "cel_79" at 972,588 size 104x54
      Appearance <- "CellSt0_30"
   IOField "io_81" at 979,595 size 90x40; FormatPattern 999
      ProcessValue <- "Cell0_30"
      Appearance <- "CellSt0_30"
   Rectangle "cel_80" at 972,648 size 104x54
      Appearance <- "CellSt0_31"
   IOField "io_82" at 979,655 size 90x40; FormatPattern 999
      ProcessValue <- "Cell0_31"
      Appearance <- "CellSt0_31"
   Rectangle "cel_81" at 972,708 size 104x54
      Appearance <- "CellSt0_32"
   IOField "io_83" at 979,715 size 90x40; FormatPattern 999
      ProcessValue <- "Cell0_32"
      Appearance <- "CellSt0_32"
   Rectangle "cel_82" at 972,768 size 104x54
      Appearance <- "CellSt0_33"
   IOField "io_84" at 979,775 size 90x40; FormatPattern 999
      ProcessValue <- "Cell0_33"
      Appearance <- "CellSt0_33"
   Rectangle "cel_83" at 972,828 size 104x54
      Appearance <- "CellSt0_34"
   IOField "io_85" at 979,835 size 90x40; FormatPattern 999
      ProcessValue <- "Cell0_34"
      Appearance <- "CellSt0_34"
   Rectangle "cel_84" at 972,888 size 104x54
      Appearance <- "CellSt0_35"
   IOField "io_86" at 979,895 size 90x40; FormatPattern 999
      ProcessValue <- "Cell0_35"
      Appearance <- "CellSt0_35"
   Rectangle "cel_85" at 1086,228 size 104x54
      Appearance <- "CellSt0_36"
   IOField "io_87" at 1093,235 size 90x40; FormatPattern 999
      ProcessValue <- "Cell0_36"
      Appearance <- "CellSt0_36"
   Rectangle "cel_86" at 1086,288 size 104x54
      Appearance <- "CellSt0_37"
   IOField "io_88" at 1093,295 size 90x40; FormatPattern 999
      ProcessValue <- "Cell0_37"
      Appearance <- "CellSt0_37"
   Rectangle "cel_87" at 1086,348 size 104x54
      Appearance <- "CellSt0_38"
   IOField "io_89" at 1093,355 size 90x40; FormatPattern 999
      ProcessValue <- "Cell0_38"
      Appearance <- "CellSt0_38"
   Rectangle "cel_88" at 1086,408 size 104x54
      Appearance <- "CellSt0_39"
   IOField "io_90" at 1093,415 size 90x40; FormatPattern 999
      ProcessValue <- "Cell0_39"
      Appearance <- "CellSt0_39"
   Rectangle "cel_89" at 1086,468 size 104x54
      Appearance <- "CellSt0_40"
   IOField "io_91" at 1093,475 size 90x40; FormatPattern 999
      ProcessValue <- "Cell0_40"
      Appearance <- "CellSt0_40"
   Rectangle "cel_90" at 1086,528 size 104x54
      Appearance <- "CellSt0_41"
   IOField "io_92" at 1093,535 size 90x40; FormatPattern 999
      ProcessValue <- "Cell0_41"
      Appearance <- "CellSt0_41"
   Rectangle "cel_91" at 1086,588 size 104x54
      Appearance <- "CellSt0_42"
   IOField "io_93" at 1093,595 size 90x40; FormatPattern 999
      ProcessValue <- "Cell0_42"
      Appearance <- "CellSt0_42"
   Rectangle "cel_92" at 1086,648 size 104x54
      Appearance <- "CellSt0_43"
   IOField "io_94" at 1093,655 size 90x40; FormatPattern 999
      ProcessValue <- "Cell0_43"
      Appearance <- "CellSt0_43"
   Rectangle "cel_93" at 1086,708 size 104x54
      Appearance <- "CellSt0_44"
   IOField "io_95" at 1093,715 size 90x40; FormatPattern 999
      ProcessValue <- "Cell0_44"
      Appearance <- "CellSt0_44"
   Rectangle "cel_94" at 1086,768 size 104x54
      Appearance <- "CellSt0_45"
   IOField "io_96" at 1093,775 size 90x40; FormatPattern 999
      ProcessValue <- "Cell0_45"
      Appearance <- "CellSt0_45"
   Rectangle "cel_95" at 1086,828 size 104x54
      Appearance <- "CellSt0_46"
   IOField "io_97" at 1093,835 size 90x40; FormatPattern 999
      ProcessValue <- "Cell0_46"
      Appearance <- "CellSt0_46"
   Rectangle "cel_96" at 1086,888 size 104x54
      Appearance <- "CellSt0_47"
   IOField "io_98" at 1093,895 size 90x40; FormatPattern 999
      ProcessValue <- "Cell0_47"
      Appearance <- "CellSt0_47"
   IOField "crn_1" at 62,188 size 100x32; FormatPattern 999
      ProcessValue <- "Carried"
      HorizontalMovement <- "CraneGX"
   Rectangle "crn_2" at 566,237 size 120x36
      VerticalMovement <- "CraneY"
   TextField "frm_6" at 1220,154 size 684x300; Text 'Text'
   TextField "txt_26" at 1232,160 size 640x28; Text 'RUČNA NAREDBA'
   TextField "txt_27" at 1232,200 size 120x34; Text 'Naredba'
   SymbolicIOField "sym_1" at 1352,200 size 240x34; TextOff '0'; TextOn '1'; TextList "TL_Cmd"
      ProcessValue <- "ManCmd"
   TextField "txt_28" at 1232,244 size 120x34; Text 'x (0-3)'
   IOField "io_99" at 1352,244 size 70x34; FormatPattern 9
      ProcessValue <- "ManX"
   TextField "txt_29" at 1440,244 size 90x34; Text 'y (0-11)'
   IOField "io_100" at 1530,244 size 70x34; FormatPattern 99
      ProcessValue <- "ManY"
   TextField "txt_30" at 1232,288 size 120x34; Text 'Bay'
   SymbolicIOField "sym_2" at 1352,288 size 240x34; TextOff '0'; TextOn '1'; TextList "TL_Bay"
      ProcessValue <- "ManBay"
   Button "btn_1" at 1640,200 size 240x122; TextOff 'IZVRŠI'
      on Press: SetBit("BtnManExec")
   TextField "txt_31" at 1232,330 size 660x22; Text 'PODIGNI/SPUSTI: lokacija dizalice. x/y/Bay: cilj pomaka.'
   TextField "txt_32" at 1232,364 size 120x32; Text 'Dizalica x'
   IOField "io_101" at 1352,364 size 50x32; FormatPattern 9
      ProcessValue <- "CraneX"
   TextField "txt_33" at 1412,364 size 30x32; Text 'y'
   IOField "io_102" at 1442,364 size 50x32; FormatPattern 99
      ProcessValue <- "CraneY"
   TextField "txt_34" at 1580,364 size 70x32; Text 'Bay'
   SymbolicIOField "sym_3" at 1650,364 size 240x32; TextOff '0'; TextOn '1'; TextList "TL_Bay"
      ProcessValue <- "CraneBay"
   TextField "txt_35" at 1232,404 size 120x32; Text 'Teret (ID)'
   IOField "io_103" at 1352,404 size 80x32; FormatPattern 999
      ProcessValue <- "Carried"
   Rectangle "lmp_1" at 1580,409 size 22x22
      Appearance <- "CraneBusy"
   TextField "txt_36" at 1606,404 size 110x32; Text 'zauzeta'
   TextField "frm_7" at 1220,462 size 684x196; Text 'Text'
   TextField "txt_37" at 1232,468 size 400x28; Text 'RAVNOTEŽA BRODA (Bay 0)'
   Rectangle "lmp_2" at 1650,472 size 22x22
      Appearance <- "BalOk"
   TextField "txt_38" at 1676,468 size 220x28; Text '|L - R| <= 5'
   TextField "txt_39" at 1232,506 size 150x32; Text 'Lijevo x0-1'
   Bar "bar_1" at 1382,508 size 400x28; MinimumValue 0; MaximumValue 24
      ProcessValue <- "BalL"
   IOField "io_104" at 1790,506 size 60x32; FormatPattern 99
      ProcessValue <- "BalL"
   TextField "txt_40" at 1232,546 size 150x32; Text 'Desno x2-3'
   Bar "bar_2" at 1382,548 size 400x28; MinimumValue 0; MaximumValue 24
      ProcessValue <- "BalR"
   IOField "io_105" at 1790,546 size 60x32; FormatPattern 99
      ProcessValue <- "BalR"
   TextField "txt_41" at 1232,590 size 150x32; Text 'Razlika L-R'
   IOField "io_106" at 1382,590 size 70x32; FormatPattern s99
      ProcessValue <- "BalDiff"
   TextField "txt_42" at 1480,590 size 110x32; Text 'Pramac'
   IOField "io_107" at 1590,590 size 60x32; FormatPattern 99
      ProcessValue <- "BalF"
   TextField "txt_43" at 1680,590 size 100x32; Text 'Krma'
   IOField "io_108" at 1780,590 size 60x32; FormatPattern 99
      ProcessValue <- "BalA"
   TextField "frm_8" at 1220,666 size 684x124; Text 'Text'
   TextField "txt_44" at 1232,672 size 400x28; Text 'NAPREDAK'
   TextField "txt_45" at 1232,706 size 90x32; Text 'Istovar'
   IOField "io_109" at 1322,706 size 52x32; FormatPattern 99
      ProcessValue <- "UDone"
   IOField "io_110" at 1380,706 size 52x32; FormatPattern 99
      ProcessValue <- "UTotal"
   TextField "txt_46" at 1460,706 size 90x32; Text 'Ukrcaj'
   IOField "io_111" at 1550,706 size 52x32; FormatPattern 99
      ProcessValue <- "LDone"
   IOField "io_112" at 1608,706 size 52x32; FormatPattern 99
      ProcessValue <- "LTotal"
   TextField "txt_47" at 1690,706 size 40x32; Text 'N'
   IOField "io_113" at 1730,706 size 60x32; FormatPattern 99
      ProcessValue <- "N"
   TextField "txt_48" at 1232,748 size 90x32; Text 'Plan #'
   IOField "io_114" at 1322,748 size 40x32; FormatPattern 9
      ProcessValue <- "PlanVariant"
   Rectangle "lmp_3" at 1400,753 size 22x22
      Appearance <- "Initialized"
   TextField "txt_49" at 1426,748 size 150x32; Text 'inicijalizirano'
   Rectangle "lmp_4" at 1590,753 size 22x22
      Appearance <- "LampDone"
   TextField "txt_50" at 1616,748 size 150x32; Text 'završeno'
   TextField "frm_9" at 1220,798 size 684x218; Text 'Text'
   TextField "txt_51" at 1232,802 size 300x24; Text 'LEGENDA ĆELIJA'
   TextField "frm_10" at 1232,832 size 45x28; Text 'Text'
   TextField "txt_52" at 1285,832 size 280x28; Text '0 prazno'
   TextField "frm_11" at 1232,876 size 45x28; Text 'Text'
   TextField "txt_53" at 1285,876 size 280x28; Text '1 zauzeto'
   TextField "frm_12" at 1232,920 size 45x28; Text 'Text'
   TextField "txt_54" at 1285,920 size 280x28; Text '2 za istovar'
   TextField "frm_13" at 1232,964 size 45x28; Text 'Text'
   TextField "txt_55" at 1285,964 size 280x28; Text '3 za ukrcaj'
   TextField "frm_14" at 1568,832 size 45x28; Text 'Text'
   TextField "txt_56" at 1621,832 size 280x28; Text '4 prebačeno'
   TextField "frm_15" at 1568,876 size 45x28; Text 'Text'
   TextField "txt_57" at 1621,876 size 280x28; Text '5 trenutni izvor'
   TextField "frm_16" at 1568,920 size 45x28; Text 'Text'
   TextField "txt_58" at 1621,920 size 280x28; Text '6 trenutni cilj'
   TextField "frm_17" at 1568,964 size 45x28; Text 'Text'
   TextField "txt_59" at 1621,964 size 280x28; Text '7 neispravan ID'

screen "Score" 1920x1080, template "Tpl"
   TextField "frm_1" at 16,154 size 900x420; Text 'Text'
   TextField "txt_1" at 28,160 size 860x28; Text 'FUNKCIJA CILJA J = 0.5*T/(N*76 s) + 0.5*M/(4N)'
   TextField "txt_2" at 330,196 size 170x30; Text 'M'
   TextField "txt_3" at 510,196 size 170x30; Text 'T [s]'
   TextField "txt_4" at 690,196 size 170x30; Text 'J'
   TextField "txt_5" at 28,234 size 300x34; Text 'M (pravilo zadatka), stvarno'
   IOField "io_1" at 330,234 size 150x34; FormatPattern 99999
      ProcessValue <- "M"
   IOField "io_2" at 510,234 size 150x34; FormatPattern 99999.9
      ProcessValue <- "T"
   IOField "io_3" at 690,234 size 150x34; FormatPattern 9.9999
      ProcessValue <- "J"
   TextField "txt_6" at 28,276 size 300x34; Text 'M (FB1 brojač, MD107)'
   IOField "io_4" at 330,276 size 150x34; FormatPattern 99999
      ProcessValue <- "MFb1"
   IOField "io_5" at 690,276 size 150x34; FormatPattern 9.9999
      ProcessValue <- "JFb1"
   TextField "txt_7" at 28,318 size 300x34; Text 'Planirani rezultat'
   IOField "io_6" at 330,318 size 150x34; FormatPattern 99999
      ProcessValue <- "PredM"
   IOField "io_7" at 510,318 size 150x34; FormatPattern 99999.9
      ProcessValue <- "PredT"
   IOField "io_8" at 690,318 size 150x34; FormatPattern 9.9999
      ProcessValue <- "PredJ"
   TextField "txt_8" at 28,372 size 860x28; Text 'OPTIMIZACIJA PLANA (FB11: pohlepni plan, zatim lokalno pretraživanje)'
   TextField "txt_9" at 28,408 size 300x34; Text 'J pohlepnog plana'
   IOField "io_9" at 328,408 size 150x34; FormatPattern 9.9999
      ProcessValue <- "PredJ0"
   TextField "txt_10" at 490,408 size 200x34; Text 'Poboljšanje [%]'
   IOField "io_10" at 690,408 size 150x34; FormatPattern 99.99
      ProcessValue <- "ImpGainPct"
   TextField "txt_11" at 28,450 size 300x34; Text 'J optimiziranog plana'
   IOField "io_11" at 328,450 size 150x34; FormatPattern 9.9999
      ProcessValue <- "PredJ"
   TextField "txt_12" at 490,450 size 200x34; Text 'Evaluacije'
   IOField "io_12" at 690,450 size 150x34; FormatPattern 99999
      ProcessValue <- "ImpEvals"
   TextField "txt_13" at 28,492 size 300x34; Text 'Donja granica J (dokazana)'
   IOField "io_13" at 328,492 size 150x34; FormatPattern 9.9999
      ProcessValue <- "LbJ"
   TextField "txt_14" at 490,492 size 200x34; Text 'Udaljenost [%]'
   IOField "io_14" at 690,492 size 150x34; FormatPattern 99.99
      ProcessValue <- "GapPct"
   TextField "txt_15" at 28,534 size 300x30; Text 'Napredak planiranja [%]'
   Bar "bar_1" at 330,536 size 360x26; MinimumValue 0; MaximumValue 100
      ProcessValue <- "PlanProgress"
   IOField "io_15" at 700,532 size 80x34; FormatPattern 999
      ProcessValue <- "PlanProgress"
   TextField "frm_2" at 932,154 size 972x420; Text 'Text'
   TextField "txt_16" at 944,160 size 940x28; Text 'POSTAVKE PLANERA'
   TextField "txt_17" at 944,200 size 260x34; Text 'Redoslijed (korišten)'
   SymbolicIOField "sym_1" at 1204,200 size 380x34; TextOff '0'; TextOn '1'; TextList "TL_Order"
      ProcessValue <- "OrderModeAct"
   TextField "txt_18" at 944,242 size 260x34; Text 'Pobjednička varijanta'
   IOField "io_16" at 1204,242 size 60x34; FormatPattern 9
      ProcessValue <- "PlanVariant"
   TextField "txt_19" at 944,284 size 260x34; Text 'N (liste)'
   IOField "io_17" at 1204,284 size 80x34; FormatPattern 99
      ProcessValue <- "N"
   Rectangle "lmp_1" at 944,333 size 22x22
      Appearance <- "Planning"
   TextField "txt_20" at 972,326 size 300x34; Text 'planiranje u tijeku'
   TextField "txt_21" at 944,380 size 940x26; Text 'Donja granica: T >= 40 s po kontejneru + 6 s po stupcu minimalnog x-puta (zatvorena formula),'
   TextField "txt_22" at 944,406 size 940x26; Text 'M >= 4 po kontejneru. Nijedan plan ne može biti bolji od te vrijednosti.'
   TextField "txt_23" at 944,442 size 940x26; Text 'Lokalno pretraživanje: premještanje, zamjena i premještanje para transfera; fiksni broj evaluacija,'
   TextField "txt_24" at 944,468 size 940x26; Text 'deterministički, uz pravilo ravnoteže |L-R| <= 5 u svakom koraku. Plan nikad nije lošiji od pohlepnog.'

screen "Screen_1" 1920x1080, template "Tpl"
   TextField "txt_1" at 60,154 size 446x28; Text 'BAY 1 - SKLADIŠTE (yard)'
   TextField "txt_2" at 744,154 size 446x28; Text 'BAY 0 - BROD (ship)'
   TextField "frm_1" at 56,186 size 1138x36; Text 'Text'
   TextField "frm_2" at 556,224 size 140x722; Text 'Text'
   TextField "txt_3" at 556,950 size 140x22; Text 'OBALA / kran y'
   TextField "frm_3" at 52,220 size 462x730; Text 'Text'
   TextField "frm_4" at 736,220 size 462x730; Text 'Text'
   TextField "frm_5" at 965,220 size 4x730; Text 'Text'
   TextField "txt_4" at 16,244 size 40x22; Text 'y0'
   TextField "txt_5" at 16,304 size 40x22; Text 'y1'
   TextField "txt_6" at 16,364 size 40x22; Text 'y2'
   TextField "txt_7" at 16,424 size 40x22; Text 'y3'
   TextField "txt_8" at 16,484 size 40x22; Text 'y4'
   TextField "txt_9" at 16,544 size 40x22; Text 'y5'
   TextField "txt_10" at 16,604 size 40x22; Text 'y6'
   TextField "txt_11" at 16,664 size 40x22; Text 'y7'
   TextField "txt_12" at 16,724 size 40x22; Text 'y8'
   TextField "txt_13" at 16,784 size 40x22; Text 'y9'
   TextField "txt_14" at 16,844 size 40x22; Text 'y10'
   TextField "txt_15" at 16,904 size 40x22; Text 'y11'
   TextField "txt_16" at 60,952 size 104x20; Text 'x0'
   TextField "txt_17" at 174,952 size 104x20; Text 'x1'
   TextField "txt_18" at 288,952 size 104x20; Text 'x2'
   TextField "txt_19" at 402,952 size 104x20; Text 'x3'
   TextField "txt_20" at 744,952 size 104x20; Text 'x0'
   TextField "txt_21" at 858,952 size 104x20; Text 'x1'
   TextField "txt_22" at 972,952 size 104x20; Text 'x2'
   TextField "txt_23" at 1086,952 size 104x20; Text 'x3'
   TextField "txt_24" at 744,976 size 120x28; Text 'LIJEVO'
   IOField "io_1" at 864,976 size 60x28; FormatPattern 99
      ProcessValue <- "BalL"
   TextField "txt_25" at 972,976 size 120x28; Text 'DESNO'
   IOField "io_2" at 1092,976 size 60x28; FormatPattern 99
      ProcessValue <- "BalR"
   Rectangle "cel_1" at 60,228 size 104x54
      Appearance <- "CellSt1_00"
   IOField "io_3" at 67,235 size 90x40; FormatPattern 999
      ProcessValue <- "Cell1_00"
      Appearance <- "CellSt1_00"
   Rectangle "cel_2" at 60,288 size 104x54
      Appearance <- "CellSt1_01"
   IOField "io_4" at 67,295 size 90x40; FormatPattern 999
      ProcessValue <- "Cell1_01"
      Appearance <- "CellSt1_01"
   Rectangle "cel_3" at 60,348 size 104x54
      Appearance <- "CellSt1_02"
   IOField "io_5" at 67,355 size 90x40; FormatPattern 999
      ProcessValue <- "Cell1_02"
      Appearance <- "CellSt1_02"
   Rectangle "cel_4" at 60,408 size 104x54
      Appearance <- "CellSt1_03"
   IOField "io_6" at 67,415 size 90x40; FormatPattern 999
      ProcessValue <- "Cell1_03"
      Appearance <- "CellSt1_03"
   Rectangle "cel_5" at 60,468 size 104x54
      Appearance <- "CellSt1_04"
   IOField "io_7" at 67,475 size 90x40; FormatPattern 999
      ProcessValue <- "Cell1_04"
      Appearance <- "CellSt1_04"
   Rectangle "cel_6" at 60,528 size 104x54
      Appearance <- "CellSt1_05"
   IOField "io_8" at 67,535 size 90x40; FormatPattern 999
      ProcessValue <- "Cell1_05"
      Appearance <- "CellSt1_05"
   Rectangle "cel_7" at 60,588 size 104x54
      Appearance <- "CellSt1_06"
   IOField "io_9" at 67,595 size 90x40; FormatPattern 999
      ProcessValue <- "Cell1_06"
      Appearance <- "CellSt1_06"
   Rectangle "cel_8" at 60,648 size 104x54
      Appearance <- "CellSt1_07"
   IOField "io_10" at 67,655 size 90x40; FormatPattern 999
      ProcessValue <- "Cell1_07"
      Appearance <- "CellSt1_07"
   Rectangle "cel_9" at 60,708 size 104x54
      Appearance <- "CellSt1_08"
   IOField "io_11" at 67,715 size 90x40; FormatPattern 999
      ProcessValue <- "Cell1_08"
      Appearance <- "CellSt1_08"
   Rectangle "cel_10" at 60,768 size 104x54
      Appearance <- "CellSt1_09"
   IOField "io_12" at 67,775 size 90x40; FormatPattern 999
      ProcessValue <- "Cell1_09"
      Appearance <- "CellSt1_09"
   Rectangle "cel_11" at 60,828 size 104x54
      Appearance <- "CellSt1_10"
   IOField "io_13" at 67,835 size 90x40; FormatPattern 999
      ProcessValue <- "Cell1_10"
      Appearance <- "CellSt1_10"
   Rectangle "cel_12" at 60,888 size 104x54
      Appearance <- "CellSt1_11"
   IOField "io_14" at 67,895 size 90x40; FormatPattern 999
      ProcessValue <- "Cell1_11"
      Appearance <- "CellSt1_11"
   Rectangle "cel_13" at 174,228 size 104x54
      Appearance <- "CellSt1_12"
   IOField "io_15" at 181,235 size 90x40; FormatPattern 999
      ProcessValue <- "Cell1_12"
      Appearance <- "CellSt1_12"
   Rectangle "cel_14" at 174,288 size 104x54
      Appearance <- "CellSt1_13"
   IOField "io_16" at 181,295 size 90x40; FormatPattern 999
      ProcessValue <- "Cell1_13"
      Appearance <- "CellSt1_13"
   Rectangle "cel_15" at 174,348 size 104x54
      Appearance <- "CellSt1_14"
   IOField "io_17" at 181,355 size 90x40; FormatPattern 999
      ProcessValue <- "Cell1_14"
      Appearance <- "CellSt1_14"
   Rectangle "cel_16" at 174,408 size 104x54
      Appearance <- "CellSt1_15"
   IOField "io_18" at 181,415 size 90x40; FormatPattern 999
      ProcessValue <- "Cell1_15"
      Appearance <- "CellSt1_15"
   Rectangle "cel_17" at 174,468 size 104x54
      Appearance <- "CellSt1_16"
   IOField "io_19" at 181,475 size 90x40; FormatPattern 999
      ProcessValue <- "Cell1_16"
      Appearance <- "CellSt1_16"
   Rectangle "cel_18" at 174,528 size 104x54
      Appearance <- "CellSt1_17"
   IOField "io_20" at 181,535 size 90x40; FormatPattern 999
      ProcessValue <- "Cell1_17"
      Appearance <- "CellSt1_17"
   Rectangle "cel_19" at 174,588 size 104x54
      Appearance <- "CellSt1_18"
   IOField "io_21" at 181,595 size 90x40; FormatPattern 999
      ProcessValue <- "Cell1_18"
      Appearance <- "CellSt1_18"
   Rectangle "cel_20" at 174,648 size 104x54
      Appearance <- "CellSt1_19"
   IOField "io_22" at 181,655 size 90x40; FormatPattern 999
      ProcessValue <- "Cell1_19"
      Appearance <- "CellSt1_19"
   Rectangle "cel_21" at 174,708 size 104x54
      Appearance <- "CellSt1_20"
   IOField "io_23" at 181,715 size 90x40; FormatPattern 999
      ProcessValue <- "Cell1_20"
      Appearance <- "CellSt1_20"
   Rectangle "cel_22" at 174,768 size 104x54
      Appearance <- "CellSt1_21"
   IOField "io_24" at 181,775 size 90x40; FormatPattern 999
      ProcessValue <- "Cell1_21"
      Appearance <- "CellSt1_21"
   Rectangle "cel_23" at 174,828 size 104x54
      Appearance <- "CellSt1_22"
   IOField "io_25" at 181,835 size 90x40; FormatPattern 999
      ProcessValue <- "Cell1_22"
      Appearance <- "CellSt1_22"
   Rectangle "cel_24" at 174,888 size 104x54
      Appearance <- "CellSt1_23"
   IOField "io_26" at 181,895 size 90x40; FormatPattern 999
      ProcessValue <- "Cell1_23"
      Appearance <- "CellSt1_23"
   Rectangle "cel_25" at 288,228 size 104x54
      Appearance <- "CellSt1_24"
   IOField "io_27" at 295,235 size 90x40; FormatPattern 999
      ProcessValue <- "Cell1_24"
      Appearance <- "CellSt1_24"
   Rectangle "cel_26" at 288,288 size 104x54
      Appearance <- "CellSt1_25"
   IOField "io_28" at 295,295 size 90x40; FormatPattern 999
      ProcessValue <- "Cell1_25"
      Appearance <- "CellSt1_25"
   Rectangle "cel_27" at 288,348 size 104x54
      Appearance <- "CellSt1_26"
   IOField "io_29" at 295,355 size 90x40; FormatPattern 999
      ProcessValue <- "Cell1_26"
      Appearance <- "CellSt1_26"
   Rectangle "cel_28" at 288,408 size 104x54
      Appearance <- "CellSt1_27"
   IOField "io_30" at 295,415 size 90x40; FormatPattern 999
      ProcessValue <- "Cell1_27"
      Appearance <- "CellSt1_27"
   Rectangle "cel_29" at 288,468 size 104x54
      Appearance <- "CellSt1_28"
   IOField "io_31" at 295,475 size 90x40; FormatPattern 999
      ProcessValue <- "Cell1_28"
      Appearance <- "CellSt1_28"
   Rectangle "cel_30" at 288,528 size 104x54
      Appearance <- "CellSt1_29"
   IOField "io_32" at 295,535 size 90x40; FormatPattern 999
      ProcessValue <- "Cell1_29"
      Appearance <- "CellSt1_29"
   Rectangle "cel_31" at 288,588 size 104x54
      Appearance <- "CellSt1_30"
   IOField "io_33" at 295,595 size 90x40; FormatPattern 999
      ProcessValue <- "Cell1_30"
      Appearance <- "CellSt1_30"
   Rectangle "cel_32" at 288,648 size 104x54
      Appearance <- "CellSt1_31"
   IOField "io_34" at 295,655 size 90x40; FormatPattern 999
      ProcessValue <- "Cell1_31"
      Appearance <- "CellSt1_31"
   Rectangle "cel_33" at 288,708 size 104x54
      Appearance <- "CellSt1_32"
   IOField "io_35" at 295,715 size 90x40; FormatPattern 999
      ProcessValue <- "Cell1_32"
      Appearance <- "CellSt1_32"
   Rectangle "cel_34" at 288,768 size 104x54
      Appearance <- "CellSt1_33"
   IOField "io_36" at 295,775 size 90x40; FormatPattern 999
      ProcessValue <- "Cell1_33"
      Appearance <- "CellSt1_33"
   Rectangle "cel_35" at 288,828 size 104x54
      Appearance <- "CellSt1_34"
   IOField "io_37" at 295,835 size 90x40; FormatPattern 999
      ProcessValue <- "Cell1_34"
      Appearance <- "CellSt1_34"
   Rectangle "cel_36" at 288,888 size 104x54
      Appearance <- "CellSt1_35"
   IOField "io_38" at 295,895 size 90x40; FormatPattern 999
      ProcessValue <- "Cell1_35"
      Appearance <- "CellSt1_35"
   Rectangle "cel_37" at 402,228 size 104x54
      Appearance <- "CellSt1_36"
   IOField "io_39" at 409,235 size 90x40; FormatPattern 999
      ProcessValue <- "Cell1_36"
      Appearance <- "CellSt1_36"
   Rectangle "cel_38" at 402,288 size 104x54
      Appearance <- "CellSt1_37"
   IOField "io_40" at 409,295 size 90x40; FormatPattern 999
      ProcessValue <- "Cell1_37"
      Appearance <- "CellSt1_37"
   Rectangle "cel_39" at 402,348 size 104x54
      Appearance <- "CellSt1_38"
   IOField "io_41" at 409,355 size 90x40; FormatPattern 999
      ProcessValue <- "Cell1_38"
      Appearance <- "CellSt1_38"
   Rectangle "cel_40" at 402,408 size 104x54
      Appearance <- "CellSt1_39"
   IOField "io_42" at 409,415 size 90x40; FormatPattern 999
      ProcessValue <- "Cell1_39"
      Appearance <- "CellSt1_39"
   Rectangle "cel_41" at 402,468 size 104x54
      Appearance <- "CellSt1_40"
   IOField "io_43" at 409,475 size 90x40; FormatPattern 999
      ProcessValue <- "Cell1_40"
      Appearance <- "CellSt1_40"
   Rectangle "cel_42" at 402,528 size 104x54
      Appearance <- "CellSt1_41"
   IOField "io_44" at 409,535 size 90x40; FormatPattern 999
      ProcessValue <- "Cell1_41"
      Appearance <- "CellSt1_41"
   Rectangle "cel_43" at 402,588 size 104x54
      Appearance <- "CellSt1_42"
   IOField "io_45" at 409,595 size 90x40; FormatPattern 999
      ProcessValue <- "Cell1_42"
      Appearance <- "CellSt1_42"
   Rectangle "cel_44" at 402,648 size 104x54
      Appearance <- "CellSt1_43"
   IOField "io_46" at 409,655 size 90x40; FormatPattern 999
      ProcessValue <- "Cell1_43"
      Appearance <- "CellSt1_43"
   Rectangle "cel_45" at 402,708 size 104x54
      Appearance <- "CellSt1_44"
   IOField "io_47" at 409,715 size 90x40; FormatPattern 999
      ProcessValue <- "Cell1_44"
      Appearance <- "CellSt1_44"
   Rectangle "cel_46" at 402,768 size 104x54
      Appearance <- "CellSt1_45"
   IOField "io_48" at 409,775 size 90x40; FormatPattern 999
      ProcessValue <- "Cell1_45"
      Appearance <- "CellSt1_45"
   Rectangle "cel_47" at 402,828 size 104x54
      Appearance <- "CellSt1_46"
   IOField "io_49" at 409,835 size 90x40; FormatPattern 999
      ProcessValue <- "Cell1_46"
      Appearance <- "CellSt1_46"
   Rectangle "cel_48" at 402,888 size 104x54
      Appearance <- "CellSt1_47"
   IOField "io_50" at 409,895 size 90x40; FormatPattern 999
      ProcessValue <- "Cell1_47"
      Appearance <- "CellSt1_47"
   Rectangle "cel_49" at 744,228 size 104x54
      Appearance <- "CellSt0_00"
   IOField "io_51" at 751,235 size 90x40; FormatPattern 999
      ProcessValue <- "Cell0_00"
      Appearance <- "CellSt0_00"
   Rectangle "cel_50" at 744,288 size 104x54
      Appearance <- "CellSt0_01"
   IOField "io_52" at 751,295 size 90x40; FormatPattern 999
      ProcessValue <- "Cell0_01"
      Appearance <- "CellSt0_01"
   Rectangle "cel_51" at 744,348 size 104x54
      Appearance <- "CellSt0_02"
   IOField "io_53" at 751,355 size 90x40; FormatPattern 999
      ProcessValue <- "Cell0_02"
      Appearance <- "CellSt0_02"
   Rectangle "cel_52" at 744,408 size 104x54
      Appearance <- "CellSt0_03"
   IOField "io_54" at 751,415 size 90x40; FormatPattern 999
      ProcessValue <- "Cell0_03"
      Appearance <- "CellSt0_03"
   Rectangle "cel_53" at 744,468 size 104x54
      Appearance <- "CellSt0_04"
   IOField "io_55" at 751,475 size 90x40; FormatPattern 999
      ProcessValue <- "Cell0_04"
      Appearance <- "CellSt0_04"
   Rectangle "cel_54" at 744,528 size 104x54
      Appearance <- "CellSt0_05"
   IOField "io_56" at 751,535 size 90x40; FormatPattern 999
      ProcessValue <- "Cell0_05"
      Appearance <- "CellSt0_05"
   Rectangle "cel_55" at 744,588 size 104x54
      Appearance <- "CellSt0_06"
   IOField "io_57" at 751,595 size 90x40; FormatPattern 999
      ProcessValue <- "Cell0_06"
      Appearance <- "CellSt0_06"
   Rectangle "cel_56" at 744,648 size 104x54
      Appearance <- "CellSt0_07"
   IOField "io_58" at 751,655 size 90x40; FormatPattern 999
      ProcessValue <- "Cell0_07"
      Appearance <- "CellSt0_07"
   Rectangle "cel_57" at 744,708 size 104x54
      Appearance <- "CellSt0_08"
   IOField "io_59" at 751,715 size 90x40; FormatPattern 999
      ProcessValue <- "Cell0_08"
      Appearance <- "CellSt0_08"
   Rectangle "cel_58" at 744,768 size 104x54
      Appearance <- "CellSt0_09"
   IOField "io_60" at 751,775 size 90x40; FormatPattern 999
      ProcessValue <- "Cell0_09"
      Appearance <- "CellSt0_09"
   Rectangle "cel_59" at 744,828 size 104x54
      Appearance <- "CellSt0_10"
   IOField "io_61" at 751,835 size 90x40; FormatPattern 999
      ProcessValue <- "Cell0_10"
      Appearance <- "CellSt0_10"
   Rectangle "cel_60" at 744,888 size 104x54
      Appearance <- "CellSt0_11"
   IOField "io_62" at 751,895 size 90x40; FormatPattern 999
      ProcessValue <- "Cell0_11"
      Appearance <- "CellSt0_11"
   Rectangle "cel_61" at 858,228 size 104x54
      Appearance <- "CellSt0_12"
   IOField "io_63" at 865,235 size 90x40; FormatPattern 999
      ProcessValue <- "Cell0_12"
      Appearance <- "CellSt0_12"
   Rectangle "cel_62" at 858,288 size 104x54
      Appearance <- "CellSt0_13"
   IOField "io_64" at 865,295 size 90x40; FormatPattern 999
      ProcessValue <- "Cell0_13"
      Appearance <- "CellSt0_13"
   Rectangle "cel_63" at 858,348 size 104x54
      Appearance <- "CellSt0_14"
   IOField "io_65" at 865,355 size 90x40; FormatPattern 999
      ProcessValue <- "Cell0_14"
      Appearance <- "CellSt0_14"
   Rectangle "cel_64" at 858,408 size 104x54
      Appearance <- "CellSt0_15"
   IOField "io_66" at 865,415 size 90x40; FormatPattern 999
      ProcessValue <- "Cell0_15"
      Appearance <- "CellSt0_15"
   Rectangle "cel_65" at 858,468 size 104x54
      Appearance <- "CellSt0_16"
   IOField "io_67" at 865,475 size 90x40; FormatPattern 999
      ProcessValue <- "Cell0_16"
      Appearance <- "CellSt0_16"
   Rectangle "cel_66" at 858,528 size 104x54
      Appearance <- "CellSt0_17"
   IOField "io_68" at 865,535 size 90x40; FormatPattern 999
      ProcessValue <- "Cell0_17"
      Appearance <- "CellSt0_17"
   Rectangle "cel_67" at 858,588 size 104x54
      Appearance <- "CellSt0_18"
   IOField "io_69" at 865,595 size 90x40; FormatPattern 999
      ProcessValue <- "Cell0_18"
      Appearance <- "CellSt0_18"
   Rectangle "cel_68" at 858,648 size 104x54
      Appearance <- "CellSt0_19"
   IOField "io_70" at 865,655 size 90x40; FormatPattern 999
      ProcessValue <- "Cell0_19"
      Appearance <- "CellSt0_19"
   Rectangle "cel_69" at 858,708 size 104x54
      Appearance <- "CellSt0_20"
   IOField "io_71" at 865,715 size 90x40; FormatPattern 999
      ProcessValue <- "Cell0_20"
      Appearance <- "CellSt0_20"
   Rectangle "cel_70" at 858,768 size 104x54
      Appearance <- "CellSt0_21"
   IOField "io_72" at 865,775 size 90x40; FormatPattern 999
      ProcessValue <- "Cell0_21"
      Appearance <- "CellSt0_21"
   Rectangle "cel_71" at 858,828 size 104x54
      Appearance <- "CellSt0_22"
   IOField "io_73" at 865,835 size 90x40; FormatPattern 999
      ProcessValue <- "Cell0_22"
      Appearance <- "CellSt0_22"
   Rectangle "cel_72" at 858,888 size 104x54
      Appearance <- "CellSt0_23"
   IOField "io_74" at 865,895 size 90x40; FormatPattern 999
      ProcessValue <- "Cell0_23"
      Appearance <- "CellSt0_23"
   Rectangle "cel_73" at 972,228 size 104x54
      Appearance <- "CellSt0_24"
   IOField "io_75" at 979,235 size 90x40; FormatPattern 999
      ProcessValue <- "Cell0_24"
      Appearance <- "CellSt0_24"
   Rectangle "cel_74" at 972,288 size 104x54
      Appearance <- "CellSt0_25"
   IOField "io_76" at 979,295 size 90x40; FormatPattern 999
      ProcessValue <- "Cell0_25"
      Appearance <- "CellSt0_25"
   Rectangle "cel_75" at 972,348 size 104x54
      Appearance <- "CellSt0_26"
   IOField "io_77" at 979,355 size 90x40; FormatPattern 999
      ProcessValue <- "Cell0_26"
      Appearance <- "CellSt0_26"
   Rectangle "cel_76" at 972,408 size 104x54
      Appearance <- "CellSt0_27"
   IOField "io_78" at 979,415 size 90x40; FormatPattern 999
      ProcessValue <- "Cell0_27"
      Appearance <- "CellSt0_27"
   Rectangle "cel_77" at 972,468 size 104x54
      Appearance <- "CellSt0_28"
   IOField "io_79" at 979,475 size 90x40; FormatPattern 999
      ProcessValue <- "Cell0_28"
      Appearance <- "CellSt0_28"
   Rectangle "cel_78" at 972,528 size 104x54
      Appearance <- "CellSt0_29"
   IOField "io_80" at 979,535 size 90x40; FormatPattern 999
      ProcessValue <- "Cell0_29"
      Appearance <- "CellSt0_29"
   Rectangle "cel_79" at 972,588 size 104x54
      Appearance <- "CellSt0_30"
   IOField "io_81" at 979,595 size 90x40; FormatPattern 999
      ProcessValue <- "Cell0_30"
      Appearance <- "CellSt0_30"
   Rectangle "cel_80" at 972,648 size 104x54
      Appearance <- "CellSt0_31"
   IOField "io_82" at 979,655 size 90x40; FormatPattern 999
      ProcessValue <- "Cell0_31"
      Appearance <- "CellSt0_31"
   Rectangle "cel_81" at 972,708 size 104x54
      Appearance <- "CellSt0_32"
   IOField "io_83" at 979,715 size 90x40; FormatPattern 999
      ProcessValue <- "Cell0_32"
      Appearance <- "CellSt0_32"
   Rectangle "cel_82" at 972,768 size 104x54
      Appearance <- "CellSt0_33"
   IOField "io_84" at 979,775 size 90x40; FormatPattern 999
      ProcessValue <- "Cell0_33"
      Appearance <- "CellSt0_33"
   Rectangle "cel_83" at 972,828 size 104x54
      Appearance <- "CellSt0_34"
   IOField "io_85" at 979,835 size 90x40; FormatPattern 999
      ProcessValue <- "Cell0_34"
      Appearance <- "CellSt0_34"
   Rectangle "cel_84" at 972,888 size 104x54
      Appearance <- "CellSt0_35"
   IOField "io_86" at 979,895 size 90x40; FormatPattern 999
      ProcessValue <- "Cell0_35"
      Appearance <- "CellSt0_35"
   Rectangle "cel_85" at 1086,228 size 104x54
      Appearance <- "CellSt0_36"
   IOField "io_87" at 1093,235 size 90x40; FormatPattern 999
      ProcessValue <- "Cell0_36"
      Appearance <- "CellSt0_36"
   Rectangle "cel_86" at 1086,288 size 104x54
      Appearance <- "CellSt0_37"
   IOField "io_88" at 1093,295 size 90x40; FormatPattern 999
      ProcessValue <- "Cell0_37"
      Appearance <- "CellSt0_37"
   Rectangle "cel_87" at 1086,348 size 104x54
      Appearance <- "CellSt0_38"
   IOField "io_89" at 1093,355 size 90x40; FormatPattern 999
      ProcessValue <- "Cell0_38"
      Appearance <- "CellSt0_38"
   Rectangle "cel_88" at 1086,408 size 104x54
      Appearance <- "CellSt0_39"
   IOField "io_90" at 1093,415 size 90x40; FormatPattern 999
      ProcessValue <- "Cell0_39"
      Appearance <- "CellSt0_39"
   Rectangle "cel_89" at 1086,468 size 104x54
      Appearance <- "CellSt0_40"
   IOField "io_91" at 1093,475 size 90x40; FormatPattern 999
      ProcessValue <- "Cell0_40"
      Appearance <- "CellSt0_40"
   Rectangle "cel_90" at 1086,528 size 104x54
      Appearance <- "CellSt0_41"
   IOField "io_92" at 1093,535 size 90x40; FormatPattern 999
      ProcessValue <- "Cell0_41"
      Appearance <- "CellSt0_41"
   Rectangle "cel_91" at 1086,588 size 104x54
      Appearance <- "CellSt0_42"
   IOField "io_93" at 1093,595 size 90x40; FormatPattern 999
      ProcessValue <- "Cell0_42"
      Appearance <- "CellSt0_42"
   Rectangle "cel_92" at 1086,648 size 104x54
      Appearance <- "CellSt0_43"
   IOField "io_94" at 1093,655 size 90x40; FormatPattern 999
      ProcessValue <- "Cell0_43"
      Appearance <- "CellSt0_43"
   Rectangle "cel_93" at 1086,708 size 104x54
      Appearance <- "CellSt0_44"
   IOField "io_95" at 1093,715 size 90x40; FormatPattern 999
      ProcessValue <- "Cell0_44"
      Appearance <- "CellSt0_44"
   Rectangle "cel_94" at 1086,768 size 104x54
      Appearance <- "CellSt0_45"
   IOField "io_96" at 1093,775 size 90x40; FormatPattern 999
      ProcessValue <- "Cell0_45"
      Appearance <- "CellSt0_45"
   Rectangle "cel_95" at 1086,828 size 104x54
      Appearance <- "CellSt0_46"
   IOField "io_97" at 1093,835 size 90x40; FormatPattern 999
      ProcessValue <- "Cell0_46"
      Appearance <- "CellSt0_46"
   Rectangle "cel_96" at 1086,888 size 104x54
      Appearance <- "CellSt0_47"
   IOField "io_98" at 1093,895 size 90x40; FormatPattern 999
      ProcessValue <- "Cell0_47"
      Appearance <- "CellSt0_47"
   IOField "crn_1" at 62,188 size 100x32; FormatPattern 999
      ProcessValue <- "Carried"
      HorizontalMovement <- "CraneGX"
   Rectangle "crn_2" at 566,237 size 120x36
      VerticalMovement <- "CraneY"
   TextField "frm_6" at 1220,154 size 684x300; Text 'Text'
   TextField "txt_26" at 1232,160 size 400x28; Text 'TRENUTNA NAREDBA'
   TextField "txt_27" at 1232,196 size 120x32; Text 'Naredba'
   SymbolicIOField "sym_1" at 1352,196 size 220x32; TextOff '0'; TextOn '1'; TextList "TL_Cmd"
      ProcessValue <- "CurCmd"
   TextField "txt_28" at 1580,196 size 70x32; Text 'Vrsta'
   SymbolicIOField "sym_2" at 1650,196 size 240x32; TextOff '0'; TextOn '1'; TextList "TL_Kind"
      ProcessValue <- "CurKind"
   TextField "txt_29" at 1232,236 size 120x32; Text 'Kontejner'
   IOField "io_99" at 1352,236 size 80x32; FormatPattern 999
      ProcessValue <- "CurId"
   TextField "txt_30" at 1580,236 size 70x32; Text 'Faza'
   SymbolicIOField "sym_3" at 1650,236 size 240x32; TextOff '0'; TextOn '1'; TextList "TL_Phase"
      ProcessValue <- "CurPhase"
   TextField "txt_31" at 1232,276 size 120x32; Text 'Cilj x'
   IOField "io_100" at 1352,276 size 50x32; FormatPattern 9
      ProcessValue <- "CurX"
   TextField "txt_32" at 1412,276 size 30x32; Text 'y'
   IOField "io_101" at 1442,276 size 50x32; FormatPattern 99
      ProcessValue <- "CurY"
   TextField "txt_33" at 1580,276 size 70x32; Text 'Bay'
   SymbolicIOField "sym_4" at 1650,276 size 240x32; TextOff '0'; TextOn '1'; TextList "TL_Bay"
      ProcessValue <- "CurBay"
   TextField "txt_34" at 1232,324 size 400x28; Text 'DIZALICA'
   TextField "txt_35" at 1232,360 size 120x32; Text 'Položaj x'
   IOField "io_102" at 1352,360 size 50x32; FormatPattern 9
      ProcessValue <- "CraneX"
   TextField "txt_36" at 1412,360 size 30x32; Text 'y'
   IOField "io_103" at 1442,360 size 50x32; FormatPattern 99
      ProcessValue <- "CraneY"
   TextField "txt_37" at 1580,360 size 70x32; Text 'Bay'
   SymbolicIOField "sym_5" at 1650,360 size 240x32; TextOff '0'; TextOn '1'; TextList "TL_Bay"
      ProcessValue <- "CraneBay"
   TextField "txt_38" at 1232,400 size 120x32; Text 'Teret (ID)'
   IOField "io_104" at 1352,400 size 80x32; FormatPattern 999
      ProcessValue <- "Carried"
   Rectangle "lmp_1" at 1580,405 size 22x22
      Appearance <- "CraneBusy"
   TextField "txt_39" at 1606,400 size 110x32; Text 'zauzeta'
   Rectangle "lmp_2" at 1720,405 size 22x22
      Appearance <- "Planning"
   TextField "txt_40" at 1746,400 size 150x32; Text 'planiranje'
   TextField "frm_7" at 1220,462 size 684x196; Text 'Text'
   TextField "txt_41" at 1232,468 size 400x28; Text 'RAVNOTEŽA BRODA (Bay 0)'
   Rectangle "lmp_3" at 1650,472 size 22x22
      Appearance <- "BalOk"
   TextField "txt_42" at 1676,468 size 220x28; Text '|L - R| <= 5'
   TextField "txt_43" at 1232,506 size 150x32; Text 'Lijevo x0-1'
   Bar "bar_1" at 1382,508 size 400x28; MinimumValue 0; MaximumValue 24
      ProcessValue <- "BalL"
   IOField "io_105" at 1790,506 size 60x32; FormatPattern 99
      ProcessValue <- "BalL"
   TextField "txt_44" at 1232,546 size 150x32; Text 'Desno x2-3'
   Bar "bar_2" at 1382,548 size 400x28; MinimumValue 0; MaximumValue 24
      ProcessValue <- "BalR"
   IOField "io_106" at 1790,546 size 60x32; FormatPattern 99
      ProcessValue <- "BalR"
   TextField "txt_45" at 1232,590 size 150x32; Text 'Razlika L-R'
   IOField "io_107" at 1382,590 size 70x32; FormatPattern s99
      ProcessValue <- "BalDiff"
   TextField "txt_46" at 1480,590 size 110x32; Text 'Pramac'
   IOField "io_108" at 1590,590 size 60x32; FormatPattern 99
      ProcessValue <- "BalF"
   TextField "txt_47" at 1680,590 size 100x32; Text 'Krma'
   IOField "io_109" at 1780,590 size 60x32; FormatPattern 99
      ProcessValue <- "BalA"
   TextField "frm_8" at 1220,666 size 684x124; Text 'Text'
   TextField "txt_48" at 1232,672 size 400x28; Text 'NAPREDAK'
   TextField "txt_49" at 1232,706 size 90x32; Text 'Istovar'
   IOField "io_110" at 1322,706 size 52x32; FormatPattern 99
      ProcessValue <- "UDone"
   IOField "io_111" at 1380,706 size 52x32; FormatPattern 99
      ProcessValue <- "UTotal"
   TextField "txt_50" at 1460,706 size 90x32; Text 'Ukrcaj'
   IOField "io_112" at 1550,706 size 52x32; FormatPattern 99
      ProcessValue <- "LDone"
   IOField "io_113" at 1608,706 size 52x32; FormatPattern 99
      ProcessValue <- "LTotal"
   TextField "txt_51" at 1690,706 size 40x32; Text 'N'
   IOField "io_114" at 1730,706 size 60x32; FormatPattern 99
      ProcessValue <- "N"
   TextField "txt_52" at 1232,748 size 90x32; Text 'Plan #'
   IOField "io_115" at 1322,748 size 40x32; FormatPattern 9
      ProcessValue <- "PlanVariant"
   Rectangle "lmp_4" at 1400,753 size 22x22
      Appearance <- "Initialized"
   TextField "txt_53" at 1426,748 size 150x32; Text 'inicijalizirano'
   Rectangle "lmp_5" at 1590,753 size 22x22
      Appearance <- "LampDone"
   TextField "txt_54" at 1616,748 size 150x32; Text 'završeno'
   TextField "frm_9" at 1220,798 size 684x218; Text 'Text'
   TextField "txt_55" at 1232,802 size 300x24; Text 'LEGENDA ĆELIJA'
   TextField "frm_10" at 1232,832 size 45x28; Text 'Text'
   TextField "txt_56" at 1285,832 size 280x28; Text '0 prazno'
   TextField "frm_11" at 1232,876 size 45x28; Text 'Text'
   TextField "txt_57" at 1285,876 size 280x28; Text '1 zauzeto'
   TextField "frm_12" at 1232,920 size 45x28; Text 'Text'
   TextField "txt_58" at 1285,920 size 280x28; Text '2 za istovar'
   TextField "frm_13" at 1232,964 size 45x28; Text 'Text'
   TextField "txt_59" at 1285,964 size 280x28; Text '3 za ukrcaj'
   TextField "frm_14" at 1568,832 size 45x28; Text 'Text'
   TextField "txt_60" at 1621,832 size 280x28; Text '4 prebačeno'
   TextField "frm_15" at 1568,876 size 45x28; Text 'Text'
   TextField "txt_61" at 1621,876 size 280x28; Text '5 trenutni izvor'
   TextField "frm_16" at 1568,920 size 45x28; Text 'Text'
   TextField "txt_62" at 1621,920 size 280x28; Text '6 trenutni cilj'
   TextField "frm_17" at 1568,964 size 45x28; Text 'Text'
   TextField "txt_63" at 1621,964 size 280x28; Text '7 neispravan ID'
*)